(* IEC 61131-3 sources: daoli-st-library/DL_Device (part 13) *)

(* ---- FB_DL_AxisEncBatteryWatch.st ---- *)
(*
    FB_DL_AxisEncBatteryWatch —— 绝对值编码器备用电池欠压监视与预警
    ------------------------------------------------------------------
    组件名称  : FB_DL_AxisEncBatteryWatch
    分类      : DL_Device / AxisHealth
    前缀      : FB_DL_
    版本      : 1.0.0
    溯源      : 借鉴点 —— 设备级粗粒度监视（AOI 粒度族）的「双阈值分型 +
                确认延时 + 锁存预警」组织方式，以及 NE107 健康分级公开条款
                （fault → eMaintenanceReq，warn → eOutOfSpec）。
                本件只借鉴**组织方式与分级语义**，判据 / 阈值 / 码位 100% 自有。
                clean-room 声明 —— 零代码行复制（来源闭源，按最严口径零接触）；
                定时与沿检测仅用 IEC 61131-3 标准库 TON / R_TRIG。
                许可证 —— 本件 MIT；来源标签 t2-6-rockwell-aoi（次源
                t2-8-ne107）仅作语义参考，不包含其任何受版权保护的实现。
    平台      : 纯 IEC 61131-3，CODESYS 3.5 / TwinCAT 3 / InoProShop / Machine Expert 通用
    作者      : 道莅代码库 · PLC编程专家（R71 构建轮 · 批 1 · 序号 3）
    ------------------------------------------------------------------
    功能说明  : 监视绝对值编码器备用电池电压 fBattV，双阈值迟滞判定：
                故障线 fFaultV（低于即电池将尽，断电将丢参考点）与预警线
                fWarnV（低于即建议更换），两线各带独立回差 fHystV 防临界抖振；
                越线须持续 tConfirm 才确认，确认后：
                预警线 → bWarn（实时位）+ bReplaceSoon（**锁存**建议更换位，
                电压回升不清除，必须 bReset 上升沿才解除 —— 电池已劣化属
                事实性结论，瞬时恢复不改判）；
                故障线 → bFault（锁存）+ 故障码。
                非有限电压（断线 / ADC 故障）→ **直接置 bFault 并锁存**
                （电池状态不明比欠压更危险，安全侧收紧，不等确认延时）。
                依赖声明：TYPE E_DL_Ne107Status（属主 I_DL_DeviceHealth.st，
                只引用不重声明，枚举全库唯一定义）；仅 Standard.library
                （TON / R_TRIG / ABS），零厂商方言。
                确认定时器 _tonWarn / _tonFault 每周期无条件调用（规则 ⑦），
                IN 为显式条件（含已确认自保持与回差释放线）。
    错误码    : 16#0002_3770 组态非法（阈值倒置 fWarnV <= fFaultV / 回差为负 /
                            回差吞没线间距 / 阈值非有限 / 幅值超域），锁存 —— 故障级
                16#0002_3771 电池电压非有限（断线 / ADC 故障），直接锁存 —— 故障级
                16#0002_3772 电池欠压越过故障线并经确认（断电将丢参考点），锁存
                            —— 故障级
                16#0002_3773 电池欠压越过预警线并经确认（建议更换）—— 信息级，
                            不置 bError（R45：预警不算故障）
                16#0002_3774 电压越出典型域 [0, 5] V（编码器电池典型域），趋势
                            参考 —— 信息级，不置 bError；不拦截照判（负电压亦
                            必然低于故障线，判定方向天然安全）
    码位总账  : 16#0002_3770 用 ｜ 16#0002_3771 用 ｜ 16#0002_3772 用 ｜
                16#0002_3773 用 ｜ 16#0002_3774 用
    状态机    : N/A —— 单相监视，无顺序状态机，无自有 ENUM / CASE 可写；
                两路确认计时由 TON 实例自持，属定时器状态而非顺序状态；
                健康出口复用既有枚举 E_DL_Ne107Status（只引用）
    边界与披露: 一 组态判据逐项点名（R272）：fWarnV / fFaultV / fHystV 全部
                   纳入非有限闸；阈值倒置（fWarnV <= fFaultV）拦截；
                   fHystV < 0 拦截；fHystV >= (fWarnV - fFaultV) 拦截（回差
                   吞没线间距时两线无迟滞带，判据恒真）；
                二 输入非有限 → 直接故障锁存（不走过闸判定集合，安全侧赋值
                   不引用本闸判定内的量，防自证循环）；
                三 失能（bEn = FALSE）语义写死（R303）：bWarn / bReplaceSoon /
                   bFault 输出全清零、bError 清零、码清零，但 _bFault /
                   _bWarnLatch 锁存位**不被失能清除**（失能是操作态，不是
                   复位），必须 bReset 上升沿才解除 —— 两者语义分离；
                四 定时器 _tonWarn / _tonFault 无论失能 / 故障 / 正常均在段 8
                   无条件调用，IN 为段 7 计算出的显式条件；
                五 阈值默认域标注：编码器备用电池典型域 0~5 V，fWarnV 默认
                   3.0 V / fFaultV 默认 2.7 V 仅为锂-二氧化锰扣式电池组的
                   常见参考值，**不构成工程承诺**，实际阈值以编码器手册为准；
                六 电压越域（0~5 V 外）只报信息级不拦截：判定方向与电压
                   单调性一致（越低越险），越域照判不产生危险侧偏差；
                七 锁存解除路径唯一：bReset 上升沿（R188，可到达、引脚可满足）；
                八 零全局变量、零 VAR_EXTERNAL、零物理地址、零数组下标、无除法。
    分工声明  : FB_DL_BrakeWearAccum（磨损累计）、FB_DL_SpindleWarmupSeq（热机
                顺控）等运动健康件互不相干；本件只做编码器备用电池电压域，
                不消费轴状态、不下发轴指令（R31 运动家族高危区纪律）。
    修订记录  : 2026-11-22 v1.0.0 首次入库（R71 构建轮 · 批 1 · 序号 3）
*)
FUNCTION_BLOCK FB_DL_AxisEncBatteryWatch
VAR_INPUT
    fBattV    : LREAL;                     (* 编码器备用电池电压，[V]，典型域 0..5 / the encoder backup battery voltage *)
    fWarnV    : LREAL := 3.0;              (* 预警阈值，[V]，须 > fFaultV（默认值为参考非承诺）/ the warn threshold, must exceed fFaultV *)
    fFaultV   : LREAL := 2.7;              (* 故障阈值，[V]，须 < fWarnV（默认值为参考非承诺）/ the fault threshold, must be under fWarnV *)
    fHystV    : LREAL := 0.1;              (* 迟滞回差带宽（两线共用独立回差量），[V]，域 [0, fWarnV - fFaultV) / the hysteresis band *)
    tConfirm  : TIME := T#2S;              (* 欠压确认延时，[ms]，须 >= T#0S / the undervoltage confirmation delay *)
    bEn       : BOOL := TRUE;              (* 使能，[标志]，FALSE 时出口清零（R303）/ the enable, FALSE clears the outlets *)
    bReset    : BOOL := FALSE;             (* 故障 / 预警复位，[标志]，上升沿唯一解除 / the reset, its rising edge is the only release *)
END_VAR
VAR_OUTPUT
    bWarn        : BOOL;                   (* 预警实时位（确认成立且未破回差线），[标志] / the live warn flag, confirmed and not released *)
    bFault       : BOOL;                   (* 故障锁存位（故障线确认或电压非有限），[标志] / the latched fault flag *)
    bReplaceSoon : BOOL;                   (* 建议更换锁存位（预警确认后保持至复位），[标志] / the latched replace-soon flag, held until reset *)
    eHealth      : E_DL_Ne107Status;       (* NE107 健康出口（fault → eMaintenanceReq，warn → eOutOfSpec）/ the NE 107 health outlet *)
    bValid       : BOOL;                   (* 出口可用，失能或锁存故障为 FALSE / the outlets usable *)
    bError       : BOOL;                   (* 故障标志，存在锁存故障时为 TRUE / the fault flag, raised while latched *)
    nErrCode     : UDINT;                  (* 错误码，0 = 正常，锁存回放 / the error id, 0 = ok, replayed from the latch *)
END_VAR
VAR
    _rtReset    : R_TRIG;                  (* 复位上升沿检测实例（无条件调用）/ the reset rising edge instance *)
    _tonWarn    : TON;                     (* 预警线确认延时实例（无条件调用）/ the warn line confirmation timer *)
    _tonFault   : TON;                     (* 故障线确认延时实例（无条件调用）/ the fault line confirmation timer *)
    _bFault     : BOOL;                    (* 故障锁存位，仅 bReset 上升沿解除 / the internal latched fault bit *)
    _bWarnLatch : BOOL;                    (* 建议更换锁存位，仅 bReset 上升沿解除 / the internal latched warn bit *)
    _nCodeLatch : UDINT;                   (* 锁存成因码，故障期回放 / the latched cause code, replayed while faulted *)
    _bCfgBad    : BOOL;                    (* 组态非法标志（逐拍重算，仅用于首次锁存）/ the configuration fault flag *)
    _bInBad     : BOOL;                    (* 电压非有限标志（逐拍重算）/ the input fault flag *)
    _bOutDom    : BOOL;                    (* 电压越典型域标志（逐拍重算，仅报信息级）/ the out-of-typical-domain flag *)
    _bRun       : BOOL;                    (* 运行许可 = 使能 且 无锁存故障 / the run permit *)
    _bWarnCond  : BOOL;                    (* 预警确认条件（含自保持与回差，送 TON）/ the warn confirmation condition *)
    _bFaultCond : BOOL;                    (* 故障确认条件（含自保持与回差，送 TON）/ the fault confirmation condition *)
END_VAR

// 段 1｜出口预置（统一出口预置，R256）/ segment 1, preset every outlet
bWarn        := FALSE;                     // 预警实时位预清零 / preset the live warn flag false
bFault       := FALSE;                     // 故障出口预清零 / preset the fault outlet false
bReplaceSoon := FALSE;                     // 建议更换出口预清零 / preset the replace-soon outlet false
eHealth      := E_DL_Ne107Status.eUnknown; // 健康出口预置未知（首拍语义）/ preset the health outlet to unknown
bValid       := FALSE;                     // 可用标志预清零 / preset the valid flag false
bError       := FALSE;                     // 故障标志预清零 / preset the error flag false
nErrCode     := 0;                         // 错误码预置无错 / preset the code to zero
_bWarnCond   := FALSE;                     // 预警条件预清零 / preset the warn condition false
_bFaultCond  := FALSE;                     // 故障条件预清零 / preset the fault condition false

// 段 2｜复位沿检测（无条件调用，规则 ⑦）/ segment 2, the reset edge instance, called unconditionally
_rtReset(CLK := bReset);                   // 每周期无条件刷新 / refreshed every scan without exception

// 段 3｜锁存解除：仅 bReset 上升沿，锁存码同步清零（唯一解除边，R188）/ segment 3, the only latch release edge
IF _rtReset.Q THEN                         // 复位上升沿 / the reset rising edge
    _bFault     := FALSE;                  // 解除故障锁存 / release the fault latch
    _bWarnLatch := FALSE;                  // 解除建议更换锁存 / release the replace-soon latch
    _nCodeLatch := 0;                      // 清锁存码（可到达的清除边）/ clear the latched code, a reachable clearing edge
END_IF

// 段 4｜组态守卫（边界一逐项点名，R272）/ segment 4, the configuration guard
_bCfgBad := (fWarnV <= fFaultV)                                          // 阈值倒置或重合（预警线必须高于故障线）/ the thresholds reversed or coincident
         OR (fHystV < 0.0)                                               // 回差为负 / a negative hysteresis
         OR (fHystV >= (fWarnV - fFaultV))                               // 回差吞没线间距 / the hysteresis swallows the line gap
         OR (fWarnV <> fWarnV) OR ((fWarnV - fWarnV) <> 0.0)             // 预警阈值非有限 / the warn threshold non finite
         OR (fFaultV <> fFaultV) OR ((fFaultV - fFaultV) <> 0.0)         // 故障阈值非有限 / the fault threshold non finite
         OR (fHystV <> fHystV) OR ((fHystV - fHystV) <> 0.0);            // 回差非有限 / the hysteresis non finite

// 段 5｜输入守卫：电压非有限即危险（状态不明 > 欠压，安全侧收紧）/ segment 5, the input guard
_bInBad := (fBattV <> fBattV) OR ((fBattV - fBattV) <> 0.0); // 电压非有限（NaN 自反判 + Inf 差值自反判，R79）/ the voltage non finite
_bOutDom := (fBattV < 0.0) OR (fBattV > 5.0);               // 电压越典型域 [0,5] V（信息级，不拦截照判）/ the voltage out of the typical domain

// 段 6｜首次成因锁存（故障期内不重推断，回放锁存码，R189）/ segment 6, the first-cause latch
IF NOT _bFault THEN                        // 未锁存时才有资格登记成因 / a cause is registered only while not latched
    IF _bCfgBad THEN                       // 组态非法（优先归因，组态是根因）/ an illegal configuration, the root cause first
        _bFault     := TRUE;               // 置故障锁存 / latch the fault
        _nCodeLatch := 16#0002_3770;       // 故障级：组态非法 / fault level: an illegal configuration
    ELSIF _bInBad THEN                     // 电压非有限（状态不明，直接锁存不等延时）/ the voltage non finite, latch at once
        _bFault     := TRUE;               // 置故障锁存 / latch the fault
        _nCodeLatch := 16#0002_3771;       // 故障级：电压非有限 / fault level: a non finite voltage
    END_IF
END_IF

// 段 7｜运行许可与确认条件计算（分支内不调用任何定时器）/ segment 7, the run permit and the conditions
_bRun := bEn AND NOT _bFault;              // 使能且无锁存故障 / enabled and not latched
IF _bRun THEN                              // 运行许可成立 / the run permit holds
    _bWarnCond  := (fBattV < fWarnV) OR (_tonWarn.Q AND NOT (fBattV > (fWarnV + fHystV)));  // 预警条件：破预警线，或已确认且未回升破回差线
    _bFaultCond := (fBattV < fFaultV) OR (_tonFault.Q AND NOT (fBattV > (fFaultV + fHystV))); // 故障条件：破故障线，或已确认且未回升破回差线
    IF _bFaultCond THEN                    // 故障线条件成立（过确认延时后锁存）/ the fault line condition holds
        IF NOT _bFault THEN                // 未锁存才登记 / register only while not latched
            IF _tonFault.Q THEN            // 故障线经确认延时 / the fault line confirmed
                _bFault     := TRUE;       // 置故障锁存 / latch the fault
                _nCodeLatch := 16#0002_3772; // 故障级：欠压越故障线 / fault level: under the fault line
            END_IF
        END_IF
    END_IF
    IF _bWarnCond AND _tonWarn.Q THEN      // 预警线经确认延时 / the warn line confirmed
        _bWarnLatch := TRUE;               // 建议更换锁存（复位才解除，边界三）/ latch the replace-soon flag
    END_IF
ELSE                                       // 失能或锁存故障 / disabled or latched
    _bWarnCond  := FALSE;                  // 条件清零，计时器随之复位 / clear the condition, the timer resets
    _bFaultCond := FALSE;                  // 条件清零 / clear the condition
END_IF

// 段 8｜定时器无条件周期调用（规则 ⑦，IN 为显式条件）/ segment 8, unconditional timer calls
_tonWarn(IN := _bWarnCond, PT := tConfirm);    // 预警确认计时，每周期无条件刷新 / the warn confirmation timer
_tonFault(IN := _bFaultCond, PT := tConfirm);  // 故障确认计时，每周期无条件刷新 / the fault confirmation timer

// 段 9｜出口映射（名实双出口同源，R191）/ segment 9, the outlet mapping
IF _bRun THEN                              // 运行许可成立（无锁存故障）/ the run permit holds, not latched
    bWarn  := _bWarnCond AND _tonWarn.Q;   // 预警实时位：运行中且确认完成 / the live warn flag, confirmed while running
    bFault := FALSE;                       // 无锁存故障，故障出口为假 / no latched fault, the outlet false
    bReplaceSoon := _bWarnLatch;           // 建议更换出口与锁存同源 / the replace-soon outlet shares its latch
    bValid := TRUE;                        // 出口可用 / the outlets usable
    IF bWarn THEN                          // 预警确认成立 / the warn confirmed
        nErrCode := 16#0002_3773;          // 信息级：建议更换（不置 bError，R45）/ info level: replace soon
        eHealth  := E_DL_Ne107Status.eOutOfSpec;   // 预警 → 超出规格 / warn, out of specification
    ELSE                                   // 无预警 / no warn
        eHealth := E_DL_Ne107Status.eOk;   // 正常 / ok
    END_IF
ELSE                                       // 失能或锁存故障（出口清零相）/ disabled or latched, the clearing phase
    IF NOT bEn THEN                        // 失能优先于故障归因（操作态，边界三）/ a disable takes precedence, an operator state
        bWarn   := FALSE;                  // 失能相出口清零（R303）/ zero the outlets while disabled
        bFault  := FALSE;                  // 出口清零（锁存保留）/ the outlet cleared, the latch kept
        bReplaceSoon := FALSE;             // 出口清零（锁存保留）/ the outlet cleared, the latch kept
        bError  := FALSE;                  // 失能不是故障 / a disabled block is not a fault
        nErrCode := 0;                     // 失能不发码 / no code while disabled
        eHealth := E_DL_Ne107Status.eCheckFunction; // 失能 → 功能检查（信号暂无效）/ disabled, function check
    ELSE                                   // 锁存故障相（失能优先级之上）/ the latched fault phase
        bFault  := TRUE;                   // 故障出口与锁存同源 / the fault outlet shares the latch
        bReplaceSoon := _bWarnLatch;       // 建议更换出口与锁存同源 / the replace-soon outlet shares its latch
        bWarn   := FALSE;                  // 故障相预警实时位清零（归并到故障出口）/ the live warn cleared in the fault phase
        bError  := TRUE;                   // 故障标志置位 / raise the fault flag
        nErrCode := _nCodeLatch;           // 回放锁存码 / replay the latched code
        eHealth := E_DL_Ne107Status.eMaintenanceReq; // 故障 → 需要维护 / maintenance required
    END_IF
END_IF
IF _bRun AND (NOT _bFault) AND _bOutDom THEN // 运行中且无锁存故障且越典型域 / running, not latched, out of domain
    IF nErrCode = 0 THEN                   // 不覆盖更高优先级码（信息级让位）/ never overrides a higher priority code
        nErrCode := 16#0002_3774;          // 信息级：电压越典型域 / info level: out of the typical domain
    END_IF
END_IF
END_FUNCTION_BLOCK

(* ---- FB_DL_BcdFieldPanelIO.st ---- *)
(*
  FB_DL_BcdFieldPanelIO  —  面板 BCD 拨码阵列采集/输出 / BCD thumbwheel field panel IO assembly
  分类 Category : DL_Device
  码位 Code     : 16#03_2_17
  段位说明      : 03_2 段低半字节 00~0F 已满（05 为历史空穴留存），R38 已进位 12/13 段，
                  本轮续用 1x 段，本件启用 17 格（R192）
  版本 Version  : 1.0.0
  来源 Source   : t2-1-lgf-converter — BCD 转换族的设备级阵列组装待挖项
  溯源 Origin   : clean-room 实现，未复制任何源码行
                  （与 FC_DL_BcdToWord / FC_DL_WordToBcd 分工：那两件是单路原子，本件是设备级阵列 IO 组装）
  功能 Function : 1) 4 位十进制拨码（16 位输入阵列）逐位消抖（FB_DL_SignalDebounce ×16）；
                  2) 消抖后按 4 bit/位组装 BCD 字 → FC_DL_BcdToWord 逐位解码 → 设定值 uSetValue；
                  3) 位码非法（半字节 > 9）持续 tInvalidTo → 故障级锁存（接线/拨码故障），bReset 解除；
                  4) 稳定值变化沿 bNewValue 单拍脉冲（内部锁存 + 单拍收口，禁同拍抹除）；
                  5) 输出路径：uDisplayVal 经 FC_DL_WordToBcd 回 BCD 字供面板灯显。
  边界 Boundary : ① 16 只消抖实例在主体首部 FOR 循环内无条件刷新（每拍必调，等效无条件域）；
                  ② 位序约定：abDigBits 下标 0 = 个位 BCD bit0，下标 4k..4k+3 = 第 k 位十进制位；
                  ③ tDebounce = T#0S 时消抖直通（消抖件原生语义，透传不钳制）；
                  ④ 组态域闸：tInvalidTo 非正按 1s 兜底（防非法组态令故障永不锁存）；
                  ⑤ 无状态机 CASE 主相（采集型 FB）：故障经锁存位承载，无跨相 TON 复用问题。
  依赖 Depends  : FB_DL_SignalDebounce（实例化 ×16）/ FC_DL_BcdToWord / FC_DL_WordToBcd（函数调用）
  码表 Error codes（本件格 03_2_17，子码步进 +0x100）:
    16#0003_0117 信息级：稳定设定值变化沿已捕获（bNewValue 拍）
    16#0003_0217 故障级：位码非法持续超 tInvalidTo（半字节 > 9，接线/拨码故障），锁存至复位
    16#0003_0317 信息级：回显 BCD 编码饱和（uDisplayVal > 9999，WordToBcd 溢出口径透传）

  修订历史 Revision :
    2026-11-19  v1.0.0  R39 首版（批次 2 · 序号 9）
*)

FUNCTION_BLOCK FB_DL_BcdFieldPanelIO
VAR_INPUT
    abDigBits  : ARRAY[0..15] OF BOOL;    // 拨码原始位输入阵列，下标 0 = 个位 bit0 / Raw digit bit inputs, index 0 = units bit0
    tDebounce  : TIME := T#20MS;          // 逐位消抖延时 [ms]，T#0S = 直通 / Per-bit debounce delay
    tInvalidTo : TIME := T#1S;            // 位码非法持续判据 [ms]，域 > 0（非法组态按 1s 兜底）/ Invalid-code persistence time
    uDisplayVal: UINT := 0;               // 面板回显十进制值 [0..9999]，越限走饱和路径 / Display value for the panel echo
    bReset     : BOOL := FALSE;           // 故障复位，上升沿生效 / Fault reset, rising edge
END_VAR
VAR_OUTPUT
    uSetValue  : UINT;                    // 稳定设定值 [0..9999]（逐位解码合成）/ Stable setpoint value
    bSetValid  : BOOL;                    // 设定值有效（无非法半字节）/ Setpoint validity flag
    anDigVal   : ARRAY[0..3] OF UINT;     // 逐位十进制值 [0..9]（故障位为垃圾值，以 bSetValid 为准）/ Per-digit decimal values
    uBcdEcho   : WORD;                    // 回显 BCD 码字（每半字节一位十进制）/ Echo BCD word for panel lamps
    bNewValue  : BOOL;                    // 稳定设定值变化沿，单拍脉冲 [-] / Stable value change edge, single-cycle pulse
    bError     : BOOL;                    // 故障锁存，仅故障级码置位，bReset 清除 [-] / Fault latch, cleared by reset
    uErrorId   : UDINT;                   // 事件码，0 = 无事件（故障级锁存回放）/ Event code, fault codes latched
END_VAR
VAR
    afbDeb     : ARRAY[0..15] OF FB_DL_SignalDebounce;  // 逐位消抖实例阵列，主体首部无条件刷新 / Per-bit debounce instances
    tonInvalid : TON;                     // 位码非法持续计时（单用途，无跨相复用）/ Invalid-code persistence timer
    rtReset    : R_TRIG;                  // 复位上升沿 / Reset rising edge
    i0         : INT;                     // 位遍历索引 [0..15]，移位量同域严格非负 / Bit loop index, also the shift amount
    _uStable   : WORD;                    // 消抖后稳定 BCD 字 / Debounced stable BCD word
    _uStablePrv: WORD;                    // 上拍稳定 BCD 字（变化沿基准）/ Previous stable BCD word, edge basis
    _bNibBad   : BOOL;                    // 本拍存在非法半字节 / Invalid nibble present this cycle
    _bInit     : BOOL := FALSE;           // 首扫标志，初值 FALSE，判据 NOT bInit（R19 范式）/ First-scan flag
    _bNewLatch : BOOL;                    // 变化沿内部锁存（单拍收口源）/ Change-edge internal latch
    _uEchoErr  : UDINT;                   // WordToBcd 回显错误码透传 / WordToBcd echo error passthrough
    _uDigErr0  : UDINT;                   // 个位 BcdToWord 错误码透传 / Units-digit decode error passthrough
    _uDigErr1  : UDINT;                   // 十位 BcdToWord 错误码透传 / Tens-digit decode error passthrough
    _uDigErr2  : UDINT;                   // 百位 BcdToWord 错误码透传 / Hundreds-digit decode error passthrough
    _uDigErr3  : UDINT;                   // 千位 BcdToWord 错误码透传 / Thousands-digit decode error passthrough
    _uInfo     : UDINT;                   // 本拍信息码，每拍重算 / Transient info code this cycle
    _uFault    : UDINT;                   // 故障码锁存寄存 / Latched fault code register
    _bFault    : BOOL;                    // 故障锁存位 / Latched fault bit
END_VAR
VAR CONSTANT
    DL_BFP_DIG_MASK : WORD := 16#000F;    // 半字节提取掩码（低 4 位）/ Nibble extraction mask
    DL_BFP_INVALID_TO_FBK : TIME := T#1S; // 非法持续判据兜底值 [ms] / Persistence-time fallback value
END_VAR

(* —— 段 0：定时器与边沿实例无条件周期刷新（R7 红线；消抖阵列在 FOR 内每拍全量刷新） —— *)
rtReset(CLK := bReset);                                         // 复位沿刷新，每拍必调
FOR i0 := 0 TO 15 DO                                            // 消抖阵列每拍全量刷新（等效无条件域）
    afbDeb[i0](bRawInput := abDigBits[i0],                      // 原始位输入
               tRiseDelay := tDebounce,                         // 上升确认延时（组态透传）
               tFallDelay := tDebounce,                         // 下降确认延时（组态透传）
               bEnable := TRUE);                                // 消抖恒使能
END_FOR
tonInvalid(IN := _bNibBad, PT := MAX(tInvalidTo, DL_BFP_INVALID_TO_FBK));   // 非法持续计时（单用途，组态兜底）

(* —— 段 1：单拍量预清零（锁存量 _uFault/_bFault/_bNewLatch/_uStablePrv 不入清单，R187①） —— *)
_uInfo := 16#0000_0000;             // 信息码每拍重算
_bNibBad := FALSE;                  // 非法半字节标志预清零
_bNewLatch := FALSE;                // 变化沿锁存预清零（组装段单点置位）
bNewValue := FALSE;                 // 变化沿出口单拍（统一出口映射）
uErrorId := 16#0000_0000;           // 事件码缺省无事件

(* —— 段 2：稳定 BCD 字组装（消抖后位 → 半字节拼接；移位量 = 下标，0..15 严格域内） —— *)
FOR i0 := 0 TO 15 DO
    IF afbDeb[i0].bStable THEN
        _uStable := _uStable OR SHL(WORD#1, i0);    // 置位（移位量归一：下标即移位量，非负）
    ELSE
        _uStable := _uStable AND NOT SHL(WORD#1, i0);   // 清位（移位量同域）
    END_IF
END_FOR

(* —— 段 3：首扫初始化（R19 唯一合法范式） —— *)
IF NOT _bInit THEN
    _uStablePrv := _uStable;        // 首扫：变化沿基准同步为当前稳定字
    _bInit := TRUE;
END_IF

(* —— 段 4：逐位 BCD 解码（FC_DL_BcdToWord 原子 ×4；非法半字节聚合） —— *)
FC_DL_BcdToWord(uBcd := _uStable AND 16#000F, uErrorId => _uDigErr0);   // 个位解码
FC_DL_BcdToWord(uBcd := SHR(_uStable, 4) AND 16#000F, uErrorId => _uDigErr1);   // 十位解码（SHR 正向移位，量归一）
FC_DL_BcdToWord(uBcd := SHR(_uStable, 8) AND 16#000F, uErrorId => _uDigErr2);   // 百位解码
FC_DL_BcdToWord(uBcd := SHR(_uStable, 12) AND 16#000F, uErrorId => _uDigErr3);  // 千位解码
IF (_uDigErr0 <> 0) OR (_uDigErr1 <> 0) OR (_uDigErr2 <> 0) OR (_uDigErr3 <> 0) THEN
    _bNibBad := TRUE;               // 本拍存在非法半字节（任一位 > 9）
END_IF
anDigVal[0] := FC_DL_BcdToWord(uBcd := _uStable AND 16#000F);           // 个位值（错误路径返回 0，安全侧）
anDigVal[1] := FC_DL_BcdToWord(uBcd := SHR(_uStable, 4) AND 16#000F);   // 十位值
anDigVal[2] := FC_DL_BcdToWord(uBcd := SHR(_uStable, 8) AND 16#000F);   // 百位值
anDigVal[3] := FC_DL_BcdToWord(uBcd := SHR(_uStable, 12) AND 16#000F);  // 千位值
uSetValue := anDigVal[0] + anDigVal[1] * 10 + anDigVal[2] * 100 + anDigVal[3] * 1000;   // 十进制合成

(* —— 段 5：故障锁存（非法持续到点才锁存，瞬时切换不误报） —— *)
IF tonInvalid.Q THEN
    _uFault := 16#0003_0217;        // 故障级：位码非法持续超限
    _bFault := TRUE;
END_IF
IF rtReset.Q THEN
    _bFault := FALSE;               // 清故障锁存位（唯一解除路径：bReset 上升沿）
    _uFault := 16#0000_0000;
END_IF

(* —— 段 6：有效性出口与变化沿（内部锁存 → 统一出口单拍，两段式收口） —— *)
bSetValid := NOT _bNibBad;          // 有效性 = 本拍无非法半字节（瞬时口径）
IF (NOT _bNibBad) AND (_uStable <> _uStablePrv) THEN
    _bNewLatch := TRUE;             // 稳定字变化：内部锁存置位（段 1 已预清零，同拍不抹）
    _uInfo := 16#0003_0117;         // 信息级：变化沿已捕获
END_IF
_uStablePrv := _uStable;            // 变化沿基准更新（段尾单点）
bNewValue := _bNewLatch;            // 出口 = 内部锁存（置位同拍不被抹）

(* —— 段 7：回显 BCD 编码（FC_DL_WordToBcd 原子，越限饱和码透传） —— *)
uBcdEcho := FC_DL_WordToBcd(uVal := uDisplayVal, uErrorId => _uEchoErr);
IF _uEchoErr <> 0 THEN
    _uInfo := 16#0003_0317;         // 信息级：回显饱和（覆盖变化沿码，回显状态优先）
END_IF

(* —— 段 8：事件码单点回放（故障锁存优先） —— *)
IF _bFault THEN
    uErrorId := _uFault;            // 故障锁存码回放
    bError := TRUE;
ELSE
    uErrorId := _uInfo;             // 信息码
    bError := FALSE;
END_IF

END_FUNCTION_BLOCK

(* ---- FB_DL_BilletShearGaugeSeq.st ---- *)
(*
  Component : FB_DL_BilletShearGaugeSeq
  Category  : DL_Device
  Type      : FB
  Complexity: C2
  VERSION   : v1.0.0
  功能      : 铸锭定尺剪切时序控制：ENUM 八态（Idle/Feed/Measure/Clamp/Shear/Trim/Release/Fault），按定尺长度送进、夹紧确认后剪切，首件去头尾。
  开源溯源  : 道莅原创 clean-room 自研（无外部代码引用）｜License: MIT
  边界条件  : ① 定尺长度须 > 1e-9、各段时长为 0 判组态非法，拒绝启动并锁存故障；
              ② 首件定尺 = 定尺长度 + 去头尾长度，去头尾仅首件执行一次；
              ③ 夹紧超时 / 松开超时均判故障，故障锁存唯一解除路径 = bReset 上升沿。
*)

TYPE E_DL_ShearPhase :
(
    eIdle    := 0,    (* 空闲：等启动沿 / Idle waiting start edge *)
    eFeed    := 10,   (* 送进：至定尺到位 / Feeding to gauge length *)
    eMeasure := 20,   (* 测长：稳定驻留 / Measuring dwell *)
    eClamp   := 30,   (* 夹紧：至夹紧反馈 / Clamping to feedback *)
    eShear   := 40,   (* 剪切：剪切保持 / Shearing hold *)
    eTrim    := 50,   (* 去头尾：首件端部切除 / Head-trim cut on first piece *)
    eRelease := 60,   (* 松开：至松开确认 / Releasing to confirmation *)
    eFault   := 90    (* 故障：锁存待复位 / Fault latched *)
);
END_TYPE

FUNCTION_BLOCK FB_DL_BilletShearGaugeSeq
VAR_INPUT
    bEnable     : BOOL;   (* 使能电平 [-] Enable level *)
    bReset      : BOOL;   (* 复位上升沿，清故障锁存 [-] Reset edge *)
    bStart      : BOOL;   (* 启动上升沿 [-] Start edge *)
    fLengthMm   : REAL;   (* 送进实测长度 [mm] Measured feed length *)
    fGaugeLenMm : REAL;   (* 定尺长度 [mm] Gauge length setpoint *)
    fTrimLenMm  : REAL;   (* 去头尾长度 [mm] Head trim length *)
    bClampFb    : BOOL;   (* 夹紧到位反馈 [-] Clamp feedback *)
    bShearFb    : BOOL;   (* 剪切到位反馈 [-] Shear feedback *)
    tMeasure    : TIME;   (* 测长驻留 [ms] Measuring dwell *)
    tShear      : TIME;   (* 剪切保持 [ms] Shear hold *)
    tTrim       : TIME;   (* 去头尾保持 [ms] Trim hold *)
    tClampTo    : TIME;   (* 夹紧超时 [ms] Clamp timeout *)
    tReleaseTo  : TIME;   (* 松开超时 [ms] Release timeout *)
END_VAR
VAR_OUTPUT
    bFeedRun    : BOOL;              (* 送进运行输出 [-] Feed run output *)
    bClampCmd   : BOOL;              (* 夹紧指令输出 [-] Clamp command *)
    bShearCmd   : BOOL;              (* 剪切指令输出 [-] Shear command *)
    bTrimCmd    : BOOL;              (* 去头尾刀指令输出 [-] Trim cut command *)
    bReleaseCmd : BOOL;              (* 松开指令输出 [-] Release command *)
    nPieceCnt   : INT;               (* 完成件数 [-] Finished piece counter *)
    ePhase      : E_DL_ShearPhase;   (* 相位出口，段尾单点映射 [-] Phase outlet *)
    bError      : BOOL;              (* 故障锁存标志 [-] Fault latch flag *)
    uErrId      : UDINT;             (* 事件码，0 = 无事件 [-] Event code *)
END_VAR
VAR
    rtReset   : R_TRIG;   (* 复位沿实例，每拍无条件刷新 / Reset edge *)
    rtStart   : R_TRIG;   (* 启动沿实例，每拍无条件刷新 / Start edge *)
    tonMeasure: TON;      (* 测长驻留计时（独立实例） / Measuring timer *)
    tonShear  : TON;      (* 剪切保持计时（独立实例） / Shear timer *)
    tonTrim   : TON;      (* 去头尾保持计时（独立实例） / Trim timer *)
    tonClampTo: TON;      (* 夹紧超时（专用超时件） / Clamp timeout *)
    tonRelTo  : TON;      (* 松开超时（专用超时件） / Release timeout *)
    _ePhase   : E_DL_ShearPhase := E_DL_ShearPhase.eIdle;  (* 内部相位 / Internal phase *)
    _bFault   : BOOL;     (* 故障锁存位（锁存量） / Latched fault bit *)
    _uFault   : UDINT;    (* 故障码锁存（锁存量） / Latched fault code *)
    _bFirst   : BOOL;     (* 首件标志（锁存量） / First piece flag *)
    _bCfgBad  : BOOL;     (* 组态非法当拍量 [-] Config illegal flag *)
    _bNonFin  : BOOL;     (* 输入非有限当拍量 [-] Non-finite input flag *)
    fTargetMm : REAL;     (* 本件定尺目标 [mm] Target length of this piece *)
END_VAR
VAR CONSTANT
    DL_EPS : REAL := 1.0E-9;   (* 浮点比较容差 [无量纲] Float compare tolerance *)
    DL_ZERO: REAL := 0.0;      (* 零常量 [-] Zero constant *)
END_VAR

(* —— 段 0｜沿与定时器每拍无条件刷新（禁置于 IF/CASE 内，使能挂 IN 引脚） —— *)
rtReset(CLK := bReset);
rtStart(CLK := bStart);
tonMeasure(IN := (_ePhase = E_DL_ShearPhase.eMeasure) AND (NOT _bFault), PT := tMeasure);
tonShear  (IN := (_ePhase = E_DL_ShearPhase.eShear)   AND (NOT _bFault), PT := tShear);
tonTrim   (IN := (_ePhase = E_DL_ShearPhase.eTrim)    AND (NOT _bFault), PT := tTrim);
tonClampTo(IN := (_ePhase = E_DL_ShearPhase.eClamp)   AND (NOT _bFault), PT := tClampTo);
tonRelTo  (IN := (_ePhase = E_DL_ShearPhase.eRelease) AND (NOT _bFault), PT := tReleaseTo);

(* —— 段 1｜每拍量预清零（锁存量 _bFault/_uFault/_bFirst/nPieceCnt 不入清单） —— *)
uErrId := 16#0000_0000;
_bCfgBad := FALSE;
_bNonFin := FALSE;

(* —— 段 2｜复位沿：故障一次性清干净，相位回空闲，首件标志复原 —— *)
IF rtReset.Q THEN
    _bFault := FALSE;
    _uFault := 16#0000_0000;
    _bFirst := TRUE;
    _ePhase := E_DL_ShearPhase.eIdle;
END_IF

(* —— 段 3｜组态闸与非有限判据（覆盖定尺长度与各段时长） —— *)
IF (fGaugeLenMm <= DL_EPS) OR (fTrimLenMm < DL_ZERO) OR (tMeasure = T#0S)
   OR (tShear = T#0S) OR (tTrim = T#0S) OR (tClampTo = T#0S) OR (tReleaseTo = T#0S) THEN
    _bCfgBad := TRUE;
END_IF
IF (fLengthMm <> fLengthMm) OR ((fLengthMm - fLengthMm) <> 0.0)
   OR (fGaugeLenMm <> fGaugeLenMm) OR ((fGaugeLenMm - fGaugeLenMm) <> 0.0)
   OR (fTrimLenMm <> fTrimLenMm) OR ((fTrimLenMm - fTrimLenMm) <> 0.0) THEN
    _bNonFin := TRUE;
END_IF

(* —— 段 4｜本件定尺目标：首件叠加去头尾长度 —— *)
IF _bFirst THEN
    fTargetMm := fGaugeLenMm + fTrimLenMm;
ELSE
    fTargetMm := fGaugeLenMm;
END_IF

(* —— 段 5｜主状态机：八态全覆盖 + ELSE 兜底 —— *)
CASE _ePhase OF
E_DL_ShearPhase.eIdle:
    bFeedRun := FALSE; bClampCmd := FALSE; bShearCmd := FALSE;
    bTrimCmd := FALSE; bReleaseCmd := FALSE;
    IF rtStart.Q AND bEnable AND (NOT _bFault) AND (NOT _bCfgBad) AND (NOT _bNonFin) THEN
        nPieceCnt := 0;
        _bFirst := TRUE;
        _ePhase := E_DL_ShearPhase.eFeed;
    ELSIF rtStart.Q AND (_bFault OR _bCfgBad OR _bNonFin) THEN
        _bFault := TRUE;                  (* 带病启动拒绝 / Reject start with bad config *)
        _uFault := 16#0024_0001;
        _ePhase := E_DL_ShearPhase.eFault;
    END_IF

E_DL_ShearPhase.eFeed:
    bFeedRun := TRUE; bClampCmd := FALSE; bShearCmd := FALSE;
    bTrimCmd := FALSE; bReleaseCmd := FALSE;
    IF _bNonFin THEN
        _bFault := TRUE; _uFault := 16#0024_0002;   (* 故障级：长度反馈非有限 *)
        _ePhase := E_DL_ShearPhase.eFault;
    ELSIF fLengthMm >= fTargetMm THEN
        _ePhase := E_DL_ShearPhase.eMeasure;        (* 迁出条件 1：定尺到位 *)
    ELSIF NOT bEnable THEN
        _ePhase := E_DL_ShearPhase.eIdle;           (* 迁出条件 2：使能撤销回安全态 *)
    END_IF

E_DL_ShearPhase.eMeasure:
    bFeedRun := FALSE; bClampCmd := FALSE; bShearCmd := FALSE;
    bTrimCmd := FALSE; bReleaseCmd := FALSE;
    IF tonMeasure.Q THEN
        _ePhase := E_DL_ShearPhase.eClamp;          (* 迁出条件 1：测长驻留完成 *)
    ELSIF NOT bEnable THEN
        _ePhase := E_DL_ShearPhase.eIdle;           (* 迁出条件 2：使能撤销 *)
    END_IF

E_DL_ShearPhase.eClamp:
    bFeedRun := FALSE; bClampCmd := TRUE; bShearCmd := FALSE;
    bTrimCmd := FALSE; bReleaseCmd := FALSE;
    IF bClampFb THEN
        _ePhase := E_DL_ShearPhase.eShear;          (* 迁出条件 1：夹紧反馈到位 *)
    ELSIF tonClampTo.Q THEN
        _bFault := TRUE; _uFault := 16#0024_0003;   (* 故障级：夹紧超时 *)
        _ePhase := E_DL_ShearPhase.eFault;
    END_IF

E_DL_ShearPhase.eShear:
    bFeedRun := FALSE; bClampCmd := TRUE; bShearCmd := TRUE;
    bTrimCmd := FALSE; bReleaseCmd := FALSE;
    IF bShearFb OR tonShear.Q THEN
        IF _bFirst THEN
            _ePhase := E_DL_ShearPhase.eTrim;       (* 首件：追加去头尾刀 *)
        ELSE
            _ePhase := E_DL_ShearPhase.eRelease;    (* 迁出条件 1：剪切到位或保持到时 *)
        END_IF
    ELSIF NOT bEnable THEN
        _ePhase := E_DL_ShearPhase.eIdle;           (* 迁出条件 2：使能撤销 *)
    END_IF

E_DL_ShearPhase.eTrim:
    bFeedRun := FALSE; bClampCmd := TRUE; bShearCmd := FALSE;
    bTrimCmd := TRUE; bReleaseCmd := FALSE;
    IF tonTrim.Q THEN
        _ePhase := E_DL_ShearPhase.eRelease;        (* 迁出条件 1：去头尾保持完成 *)
    ELSIF NOT bEnable THEN
        _ePhase := E_DL_ShearPhase.eIdle;           (* 迁出条件 2：使能撤销 *)
    END_IF

E_DL_ShearPhase.eRelease:
    bFeedRun := FALSE; bClampCmd := FALSE; bShearCmd := FALSE;
    bTrimCmd := FALSE; bReleaseCmd := TRUE;
    IF NOT bClampFb THEN
        nPieceCnt := nPieceCnt + 1;                 (* 完成件数累加：仅在迁出拍执行一次 *)
        _bFirst := FALSE;                           (* 首件完成，后续按纯定尺 *)
        _ePhase := E_DL_ShearPhase.eFeed;           (* 迁出条件 1：松开确认到位 *)
    ELSIF tonRelTo.Q THEN
        _bFault := TRUE; _uFault := 16#0024_0004;   (* 故障级：松开超时 *)
        _ePhase := E_DL_ShearPhase.eFault;
    END_IF

E_DL_ShearPhase.eFault:
    bFeedRun := FALSE; bClampCmd := FALSE; bShearCmd := FALSE;
    bTrimCmd := FALSE; bReleaseCmd := FALSE;        (* 故障相：全部输出走安全侧 *)

ELSE
    _bFault := TRUE;                                (* 兜底：非法相位锁存 *)
    _uFault := 16#0024_0009;
    _ePhase := E_DL_ShearPhase.eFault;
END_CASE

(* —— 段 6｜相位与故障码出口单点映射 —— *)
ePhase := _ePhase;
bError := _bFault;
IF _bFault AND (_uFault <> 16#0000_0000) THEN
    uErrId := _uFault;                              (* 故障码锁存回放 / Latched fault replay *)
END_IF
END_FUNCTION_BLOCK

(* ---- FB_DL_BmsPdiGateway.st ---- *)
(*
  FB_DL_BmsPdiGateway  —  楼宇侧 PDI 对象网关轮询（调度 + 异常上报） / Building-side PDI object gateway polling: scheduling plus exception report
  分类 Category : DL_Device
  版本 Version  : 1.0.0
  来源 Source   : t1-4-codesys-forge — 网关轮询族零检索深化（与 PdiReadScheduler 调度底座分工：那件为底层调度，本件为楼宇网关应用件）
  溯源 Origin   : clean-room 实现，未复制任何源码行
  功能 Function : 1) 轮询调度：bPollTick 调用方节拍沿驱动，对象索引 0..uObjCnt-1
                  轮转（uObjCnt 域闸 1..8），每拍采信当前对象 bPollOk / fObjVal
                  契约快照，逐对象连续失败计数 auFailCnt；
                  2) 异常上报：连续失败达 uFailTo → 0528 首出对象锁存
                  （nFirstFailObj 记首出号，R190 归因唯一）；对象值非有限
                  → 0529 防御锁存（NaN 自反判）；
                  3) 成功承载：失败计数清零 + 值快照写入 afObjVal + 信息级
                  042E；首出锁存拍发 042F；
                  4) 故障级：0528 对象连续失败超阈 / 0529 对象值非有限 /
                  052A 组态非法（对象数越域）+ ELSE 兜底归并；
                  5) 信息级三码：轮询成功 / 超时上报 / 网关复位（单拍沿）；
                  6) 解除式全当拍量（R240 落地），逐 BOOL 标注见段 4。
  边界 Boundary : ① 分段理由（R192）：段 0003 故障带 03A0~03FF 于 R42 用尽，
                  启用 05xx 副带续编，避开 0590~0599 判错位段；
                  ② 组态闸：uObjCnt = 0 或 > 8 或 uFailTo = 0 → 052A 锁存，
                  轮询停发；对象索引域 0..7 由 uObjCnt 域闸与常量 8 结构性限定；
                  ③ 失败计数 USINT 饱和前置判（防回绕）；
                  ④ 无 GVL 依赖：纯引脚输入输出，无外部变量引用，无物理 IO 地址。
  依赖 Depends  : Standard.library（R_TRIG）
  码表 Error codes（Device 段 0003，窗口 0528~052A / 042E~0430）:
    16#0003_0528 故障级：对象连续失败超阈锁存（首出对象号入 nFirstFailObj），锁存至 bReset
    16#0003_0529 故障级：对象值非有限锁存（防御兜底），锁存至 bReset
    16#0003_052A 故障级：组态非法（对象数/失败阈域非法）或相位落 ELSE 兜底（归并声明），锁存至 bReset
    16#0003_042E 信息级：轮询成功沿（对象值快照写入拍）
    16#0003_042F 信息级：超时上报沿（首出锁存拍）
    16#0003_0430 信息级：网关复位沿（台账清零拍）
  修订历史 Revision :
    2026-11-19  v1.0.0  R42 首版（批次 4 · 序号 5）
*)

TYPE E_DL_BpgState :
(
    eIdle  := 0,     // 未使能：不轮询 / Idle, not polling
    ePoll  := 10,    // 轮询中：逐对象承载 / Poll, per-object engaged
    eFault := 90     // 故障：首出或非有限锁定 / Fault, latched
);
END_TYPE

FUNCTION_BLOCK FB_DL_BmsPdiGateway
VAR_INPUT
    bPollTick    : BOOL := FALSE;     // 轮询节拍沿（调用方驱动）[-] / Poll tick edge from caller
    bPollOk      : BOOL := FALSE;     // 当前对象轮询成功（当拍量契约）[-] / Current-object poll success
    fObjVal      : REAL := 0.0;       // 当前对象值 [工程单位]，bPollOk 当拍采信 / Current-object value
    uObjCnt      : USINT := 8;        // 对象总数 [1..8]，域闸 / Object count
    uFailTo      : USINT := 3;        // 连续失败阈 [次]，域 > 0 / Consecutive-fail threshold
    bGwEn        : BOOL := FALSE;     // 网关使能（电平）[-] / Gateway enable, level
    bReset       : BOOL := FALSE;     // 复位，上升沿清故障锁存与台账 / Reset edge
END_VAR
VAR_OUTPUT
    eState       : E_DL_BpgState;     // 状态出口，段尾单点映射 / State outlet
    nObjIdx      : DINT;              // 当前轮询对象号 [0..7]，-1 = 未轮询 / Current polling object index
    afObjVal     : ARRAY[0..7] OF REAL;   // 逐对象值快照 [工程单位] / Per-object value snapshots
    auFailCnt    : ARRAY[0..7] OF USINT;  // 逐对象连续失败计数 [次] / Per-object fail counts
    nFirstFailObj: DINT;              // 首出失败对象号 [0..7]，-1 = 无首出 / First failed object index
    bError       : BOOL;              // 故障锁存标志 / Fault latch flag
    nErrId       : UDINT;             // 事件码，0 = 无事件 / Event code
END_VAR
VAR
    rtPollTick   : R_TRIG;            // 轮询节拍沿实例，无条件刷新 / Poll tick edge instance
    rtReset      : R_TRIG;            // 复位沿实例，无条件刷新 / Reset edge instance
    _eState      : E_DL_BpgState := E_DL_BpgState.eIdle;  // 内部相位（CASE 唯一写入目标）/ Internal phase
    _nObjCursor  : UDINT := 0;        // 轮转游标 [0..uObjCnt-1] / Round-robin cursor
    _nIdx        : DINT;              // 阵列循环索引 [-] / Array loop index
    _bValNonFin  : BOOL;              // 对象值非有限当拍量 [-] / Object-value non-finite flag
    _bFault      : BOOL;              // 故障锁存位（锁存量）/ Latched fault bit
    _uFault      : UDINT;             // 故障码锁存（锁存量）/ Latched fault code
    _uInfo       : UDINT;             // 信息码，每拍重算 / Transient info code
END_VAR

(* —— 段 0：沿实例无条件周期刷新（禁置于 IF/CASE 内） —— *)
_bValNonFin := (fObjVal <> fObjVal)
            OR ((fObjVal - fObjVal) <> (fObjVal - fObjVal));    // 值非有限防御（NaN 自反 + 差值自减）
rtPollTick(CLK := bPollTick);       // 轮询节拍沿（每拍必调）
rtReset(CLK := bReset);             // 复位沿（每拍必调）

(* —— 段 1：单拍量预清零（锁存量 _bFault/_uFault 与计数阵列不入清单，禁同拍抹除） —— *)
_uInfo := 16#0000_0000;             // 信息码每拍重算
nObjIdx := -1;                      // 对象号缺省 -1
nErrId := 16#0000_0000;             // 事件码缺省无事件

(* —— 段 2：复位沿 + 组态域闸（判据当拍量） —— *)
IF rtReset.Q THEN                   // rtReset.Q = 当拍量
    _bFault := FALSE;               // 清故障锁存位
    _uFault := 16#0000_0000;        // 清故障锁存码
    nFirstFailObj := -1;            // 首出对象号恢复哨兵
    FOR _nIdx := 0 TO 7 DO          // 台账逐对象清零
        auFailCnt[_nIdx] := 0;      // 失败计数清零
        afObjVal[_nIdx] := 0.0;     // 值快照清零
    END_FOR
    _uInfo := 16#0003_0430;         // 信息级：网关复位沿
END_IF
IF (uObjCnt < 1) OR (uObjCnt > 8) OR (uFailTo = 0) THEN      // 域闸（1..8 与失败阈）
    _uFault := 16#0003_052A;        // 故障级：组态非法
    _bFault := TRUE;                // 故障标志与码位配对（R45）
END_IF

(* —— 段 3：轮询沿承载（判据当拍量；对象索引由域闸 1..8 结构性限域） —— *)
IF rtPollTick.Q AND (_eState = E_DL_BpgState.ePoll) AND (NOT _bFault) THEN
    _nObjCursor := (_nObjCursor + 1) MOD UDINT(uObjCnt);    // 轮转游标（模基数域闸 > 0，无除零）
    nObjIdx := UDINT_TO_DINT(_nObjCursor);          // 当前对象号（域 0..uObjCnt-1 ⊆ 0..7）
    IF bPollOk THEN                 // 成功承载（当拍量契约）
        auFailCnt[nObjIdx] := 0;    // 失败计数清零
        IF NOT _bValNonFin THEN     // 值快照仅非有限闸通过后写入（FB32-7 保持槽闸）
            afObjVal[nObjIdx] := fObjVal;       // 值快照写入
        END_IF
        _uInfo := 16#0003_042E;     // 信息级：轮询成功沿
    ELSE                            // 失败承载
        IF auFailCnt[nObjIdx] < 255 THEN
            auFailCnt[nObjIdx] := auFailCnt[nObjIdx] + 1;   // 计数递增（饱和前置判防回绕）
        END_IF
        IF (auFailCnt[nObjIdx] >= uFailTo) AND (nFirstFailObj = -1) THEN
            nFirstFailObj := nObjIdx;   // 首出对象号锁定（仅首个写入）
            _uFault := 16#0003_0528;    // 故障级：连续失败超阈
            _bFault := TRUE;
            _uInfo := 16#0003_042F;     // 信息级：超时上报沿
        END_IF
    END_IF
    IF _bValNonFin AND bPollOk THEN // 成功契约但值非有限：防御锁存（0529 独立归因）
        _uFault := 16#0003_0529;    // 故障级：对象值非有限
        _bFault := TRUE;
    END_IF
END_IF

(* —— 段 4：故障解除式（R240 落地，逐 BOOL 标注）：
     rtReset.Q = 当拍量；bPollOk = 当拍量；NOT bGwEn = 当拍量。
     均不含锁存量（_bFault/_uFault），解除边真实可达（轮询恢复 + 撤使能 + 复位沿）。 —— *)
IF rtReset.Q AND bPollOk AND (NOT bGwEn) THEN
    _bFault := FALSE;               // 清故障锁存位（锁存量，仅此当拍量解除沿可清）
    _uFault := 16#0000_0000;        // 清故障锁存码（锁存量，仅本当拍量解除沿可清）
    IF _eState = E_DL_BpgState.eFault THEN
        _eState := E_DL_BpgState.eIdle;     // 故障相迁出：回未使能
    END_IF
END_IF

(* —— 段 5：相位机（CASE 全覆盖 + ELSE 兜底） —— *)
CASE _eState OF

E_DL_BpgState.eIdle:
    IF bGwEn AND (NOT _bFault) THEN
        _eState := E_DL_BpgState.ePoll;     // 使能：进轮询相
    END_IF

E_DL_BpgState.ePoll:
    IF (NOT _bFault) AND (NOT bGwEn) THEN
        _eState := E_DL_BpgState.eIdle;     // 撤使能：回未使能相
    END_IF
    (* 首出/非有限迁出在段 3 承载（置 _bFault 后次拍迁故障相） *)

E_DL_BpgState.eFault:
    ;                               // 故障相：轮询冻结，等解除沿（段 4 承载迁出）

ELSE
    _uFault := 16#0003_052A;        // 故障级：非法相位兜底（归并组态码，码表声明）
    _bFault := TRUE;
    _eState := E_DL_BpgState.eFault;    // 强制回故障相

END_CASE

(* —— 段 6：出口单点映射（名实同源；锁存码回放，禁同拍抹除） —— *)
IF _bFault THEN
    nErrId := _uFault;              // 故障锁存码回放
    nObjIdx := -1;                  // 故障相对象号恢复未轮询哨兵
ELSE
    nErrId := _uInfo;               // 信息码
END_IF
bError := _bFault;                  // 故障标志与锁存位同源
eState := _eState;                  // 状态出口单点映射

END_FUNCTION_BLOCK

(* ---- FB_DL_BoilerFlueCondenseGuard.st ---- *)
(*
  FB_DL_BoilerFlueCondenseGuard  —  锅炉烟气冷凝防护（排烟温度低限联锁 + 回水温度钳制） / Boiler flue-gas condensation guard with low flue-temperature interlock and return-water clamping
  分类 Category : DL_Device
  版本 Version  : 1.0.0
  来源 Source   : t1-2-oscat-building — 楼宇锅炉防冷凝保护族深化
  溯源 Origin   : 道莅 clean-room 实现；排烟温度低限联锁 + 回水温度低限钳制为公开锅炉防低温腐蚀保护逻辑，未复制任何源码行
  功能 Function : 1) 三级判据：排烟温度 fFlueTempC 低于报警限 fFlueLoC → 冷凝风险信息位；
                  低于联锁限 fFlueLoLoC 且持续 tConfirm → 联锁撤销燃烧器许可；
                  2) 回水温度钳制：fReturnTempC 低于 fReturnMinC 时输出 bReturnClamp 请求（提高回水），
                  仅在燃烧器许可有效时给出；
                  3) 故障级单码 052C / 信息级 0432 = 冷凝风险进入沿（由无风险转风险单拍）。
  接口 Interface: 输入排烟温度/两级限值/回水温度/回水下限/确认延时；输出许可与风险位
  边界 Boundary : ① 组态闸：fFlueLoLoC >= fFlueLoC（联锁限须低于报警限）、fFlueLoC <= 0.0、
                  fReturnMinC < 0.0、tConfirm <= T#0S → 052C 锁存；
                  ② 温度非有限（NaN 自反 + Inf 差值自减）→ 052C 锁存，燃烧器许可撤销（安全侧）；
                  ③ 低限判据为「<=」单侧直比（限值语义明确，无容差歧义），回水钳制同为单侧直比；
                  ④ 一个 TON + 两个 R_TRIG 段 0 无条件调用；⑤ 故障相迁出唯一路径 = bReset 上升沿；
                  ⑥ 零全局耦合：无 GVL / VAR_EXTERNAL / %I %Q %M 直接地址。
  依赖 Depends  : Standard.library（TON / R_TRIG）
  码表 Error codes（Device 分段见下，故障窗口 052C / 信息窗口 0432）:
    16#0003_052C 故障级：烟气冷凝防护故障总码（组态非法 / 温度非有限），锁存至 bReset 上升沿；
                 归因见 eCause，不新增码位（派单硬约束单码）
    16#0003_0432 信息级：冷凝风险进入沿（无风险 → 风险，单拍）
    分段理由：段 0003 故障带 03A0~03FF 于 R42 用尽，启用 05xx 副带续编，避开 0590~0599 判错位段。
  修订历史 Revision :
    2026-11-19  v1.0.0  R43 首版（批次 4 · 序号 16）
*)

TYPE E_DL_BfgState :
(
    eIdle     := 0,   // 未使能：许可撤销 / Idle, permit withdrawn
    eGuard    := 10,  // 防护监视中（许可有效） / Guarding with permit valid
    eLockout  := 20,  // 联锁动作（许可撤销） / Interlocked, permit withdrawn
    eFault    := 90   // 故障锁存相 / Fault latched phase
);
END_TYPE

TYPE E_DL_BfgCause :
(
    eNone       := 0, // 无故障成因 / No cause
    eCfgIllegal := 1, // 组态非法 / Illegal configuration
    eNonFinite  := 2  // 温度非有限 / Non-finite temperature
);
END_TYPE

FUNCTION_BLOCK FB_DL_BoilerFlueCondenseGuard
VAR_INPUT
    fFlueTempC   : REAL := 0.0;        // 排烟温度 [°C] / Flue gas temperature
    fFlueLoC     : REAL := 90.0;       // 冷凝风险报警限 [°C]，域 > 0 / Condensation alarm limit
    fFlueLoLoC   : REAL := 70.0;       // 联锁限 [°C]，须低于报警限 / Interlock limit
    fReturnTempC : REAL := 0.0;        // 回水温度 [°C] / Return water temperature
    fReturnMinC  : REAL := 55.0;       // 回水温度下限 [°C]，域 >= 0 / Return water minimum
    tConfirm     : TIME := T#30S;      // 联锁确认延时 [ms]，域 > 0 / Interlock confirmation delay
    bEnable      : BOOL := FALSE;      // 防护使能（电平）[-] / Guard enable
    bReset       : BOOL := FALSE;      // 复位命令，上升沿清故障 [-] / Reset edge
END_VAR
VAR_OUTPUT
    eState       : E_DL_BfgState;      // 状态出口，段 6 单点映射 / State outlet
    eCause       : E_DL_BfgCause;      // 故障成因出口（R190） / Fault cause outlet
    bBurnerPermit: BOOL;               // 燃烧器许可 [-] / Burner permit
    bCondenseRisk: BOOL;               // 冷凝风险位 [-] / Condensation risk flag
    bReturnClamp : BOOL;               // 回水温度钳制请求 [-] / Return-water clamping request
    bError       : BOOL;               // 故障锁存标志 [-] / Fault latch flag
    nErrId       : UDINT;              // 事件码，0 = 无事件 / Event code
END_VAR
VAR
    _eState      : E_DL_BfgState := E_DL_BfgState.eIdle;   // 内部相位（CASE 唯一写入目标） / Internal phase
    _eCause      : E_DL_BfgCause := E_DL_BfgCause.eNone;   // 故障成因锁存（锁存量） / Latched cause
    tonConfirm   : TON;                // 联锁确认计时，每周期无条件调用 / Confirmation timer
    rtReset      : R_TRIG;             // 复位沿实例，每周期无条件调用 / Reset edge
    rtRisk       : R_TRIG;             // 风险沿实例，每周期无条件调用 / Risk edge
    _bRisk       : BOOL;               // 冷凝风险当拍量 [-] / Risk verdict
    _bLoLo       : BOOL;               // 低于联锁限当拍量 [-] / Below interlock limit
    _bRetLow     : BOOL;               // 回水低于下限当拍量 [-] / Return water below minimum
    _bNonFin     : BOOL;               // 温度非有限当拍量 [-] / Non-finite temperature
    _bCfgBad     : BOOL;               // 组态非法当拍量 [-] / Config illegal
    _bFault      : BOOL;               // 故障锁存位（锁存量） / Latched fault bit
    _uFault      : UDINT;              // 故障码锁存（锁存量） / Latched fault code
    _uInfo       : UDINT;              // 信息码，每拍重算 / Transient info code
END_VAR

(* —— 段 0：沿实例与定时器无条件周期刷新 + 当拍量判据 —— *)
_bRisk := fFlueTempC <= fFlueLoC;                                            // 冷凝风险（单侧直比） / Risk verdict
_bLoLo := fFlueTempC <= fFlueLoLoC;                                          // 低于联锁限 / Below interlock
_bRetLow := fReturnTempC < fReturnMinC;                                      // 回水低于下限 / Return below minimum
_bNonFin := (fFlueTempC <> fFlueTempC) OR (fReturnTempC <> fReturnTempC)
         OR ((fFlueTempC - fFlueTempC) <> (fFlueTempC - fFlueTempC))
         OR ((fReturnTempC - fReturnTempC) <> (fReturnTempC - fReturnTempC));  // NaN 自反 + Inf 差值自减 / NaN and Inf
_bCfgBad := (fFlueLoLoC >= fFlueLoC) OR (fFlueLoC <= 0.0) OR (fReturnMinC < 0.0)
            OR (tConfirm <= T#0S);                                           // 组态非法当拍量 / Config illegal
rtReset(CLK := bReset);                                                      // 复位沿，每拍必调 / Reset edge
rtRisk(CLK := _bRisk AND (NOT _bFault));                                     // 风险沿（故障相屏蔽） / Risk edge
tonConfirm(IN := (_eState = E_DL_BfgState.eGuard) AND _bLoLo, PT := tConfirm);   // 联锁确认计时 / Interlock timer

(* —— 段 1：单拍量预清零（锁存量不入清单） —— *)
_uInfo := 16#0000_0000;            // 信息码每拍重算 / Info recomputed
bBurnerPermit := FALSE;            // 许可缺省撤销（安全侧缺省） / Permit default withdrawn
bCondenseRisk := FALSE;            // 风险位缺省 FALSE / Risk default
bReturnClamp := FALSE;             // 钳制请求缺省 FALSE / Clamp default
nErrId := 16#0000_0000;            // 事件码缺省无事件 / Event code default

(* —— 段 2：复位沿 + 组态域闸 —— *)
IF rtReset.Q THEN                              // rtReset.Q = 当拍量 / current scan
    _bFault := FALSE;                          // 清故障锁存位（锁存量） / Clear fault latch
    _uFault := 16#0000_0000;                   // 清故障锁存码（锁存量） / Clear fault code
    _eCause := E_DL_BfgCause.eNone;            // 清成因（锁存量） / Clear cause
    IF _eState = E_DL_BfgState.eFault THEN
        _eState := E_DL_BfgState.eIdle;        // 故障相迁出：回未使能 / Fault exit to idle
    END_IF
    IF _eState = E_DL_BfgState.eLockout THEN
        _eState := E_DL_BfgState.eGuard;       // 联锁相复位迁出：回防护（恢复许可） / Lockout exit to guard
    END_IF
END_IF
IF _bCfgBad THEN                               // 组态域闸 / Config gate
    _uFault := 16#0003_052C;                   // 故障级：防护故障总码（05xx 副带） / Device fault code
    _eCause := E_DL_BfgCause.eCfgIllegal;      // 归因：组态非法 / Cause: illegal config
    _bFault := TRUE;                           // 标志与码位配对（R45） / Flag paired with code
END_IF
IF (NOT _bFault) AND _bNonFin THEN             // 非有限锁存 / Non-finite latch
    _uFault := 16#0003_052C;
    _eCause := E_DL_BfgCause.eNonFinite;       // 归因：非有限 / Cause: non-finite
    _bFault := TRUE;
END_IF

(* —— 段 3：联锁确认（低于联锁限持续 tConfirm 即进联锁相） —— *)
IF (NOT _bFault) AND (_eState = E_DL_BfgState.eGuard) AND tonConfirm.Q THEN
    _eState := E_DL_BfgState.eLockout;         // 进联锁相（许可撤销） / Enter lockout
END_IF

(* —— 段 4：故障解除式（R240；全当拍量）：rtReset.Q / NOT _bCfgBad / NOT _bNonFin —— *)
IF rtReset.Q AND (NOT _bCfgBad) AND (NOT _bNonFin) THEN
    _bFault := FALSE;                          // 清故障锁存位（锁存量） / Clear fault latch
    _uFault := 16#0000_0000;                   // 清故障锁存码（锁存量） / Clear fault code
    _eCause := E_DL_BfgCause.eNone;            // 清成因（锁存量） / Clear cause
END_IF

(* —— 段 4A：故障锁存相位迁移闸 —— *)
IF _bFault AND (_eState <> E_DL_BfgState.eFault) THEN
    _eState := E_DL_BfgState.eFault;           // 锁存即入故障相 / Latch enters fault phase
END_IF

(* —— 段 5：相位机（CASE 全覆盖 + ELSE 兜底） —— *)
CASE _eState OF

E_DL_BfgState.eIdle:
    IF bEnable AND (NOT _bFault) THEN          // 使能条件 / Enable gate
        _eState := E_DL_BfgState.eGuard;       // 进防护相 / Enter guard
    END_IF

E_DL_BfgState.eGuard:
    bBurnerPermit := NOT _bLoLo;               // 许可：未低于联锁限即允许 / Permit unless below interlock
    bCondenseRisk := _bRisk;                   // 风险位（相内按当拍量给出） / Risk flag
    bReturnClamp := _bRetLow AND bBurnerPermit; // 回水钳制请求（许可有效时） / Return clamp request
    IF rtRisk.Q THEN                           // 风险进入沿 / Risk entrance edge
        _uInfo := 16#0003_0432;                // 信息级：冷凝风险进入沿 / Info: risk entrance
    END_IF
    IF NOT bEnable THEN                        // 撤使能：许可撤销，回未使能 / Disable withdraws permit
        _eState := E_DL_BfgState.eIdle;
    ELSIF NOT _bRisk THEN                      // 风险消失：保持防护相（不迁移） / Risk cleared, stay
        ;
    END_IF

E_DL_BfgState.eLockout:
    bBurnerPermit := FALSE;                    // 联锁相：许可强制撤销 / Permit forced withdrawn
    bCondenseRisk := TRUE;                     // 联锁相风险位恒真 / Risk latched high
    IF NOT _bLoLo THEN                         // 排烟温度回到联锁限之上（事件） / Flue temperature recovered
        _eState := E_DL_BfgState.eGuard;       // 恢复防护相 / Back to guard
    ELSIF NOT bEnable THEN                     // 撤使能：回未使能 / Disable returns idle
        _eState := E_DL_BfgState.eIdle;
    END_IF

E_DL_BfgState.eFault:
    ;                                          // 故障相：许可撤销，仅段 4 复位沿可迁出 / Permit withdrawn, reset only

ELSE
    _uFault := 16#0003_052C;                   // 故障级：非法相位兜底（归并总码） / Illegal phase fallback
    _eCause := E_DL_BfgCause.eCfgIllegal;      // 归因：相位非法归并组态 / Cause: phase illegal
    _bFault := TRUE;
    _eState := E_DL_BfgState.eFault;           // 强制回故障相 / Force fault phase

END_CASE

(* —— 段 6：出口单点映射（名实同源；故障相许可强制撤销） —— *)
IF _bFault THEN
    bBurnerPermit := FALSE;                    // 故障相许可强制撤销（安全侧） / Permit forced withdrawn
    bReturnClamp := FALSE;                     // 故障相钳制请求强制 FALSE / Clamp forced false
    nErrId := _uFault;                         // 故障锁存码回放 / Replay latched code
ELSE
    nErrId := _uInfo;                          // 信息码 / Transient info
END_IF
bError := _bFault;                             // 故障标志同源 / Flag from latch
eState := _eState;                             // 状态出口 / State outlet
eCause := _eCause;                             // 成因出口 / Cause outlet

END_FUNCTION_BLOCK

(* ---- FB_DL_BoothExhaustDamperSeq.st ---- *)
(*
  Name: FB_DL_BoothExhaustDamperSeq
  Category: DL_Device
  Version: 1.0.0
  Round: R89 / 2026-11-25
  开源溯源：clean-room 自研（族 涂装喷涂线，ST 开源生态实测 0 命中，无外部代码引入）
  功能：喷房排风风门开度顺序：起机预吹→生产→清洗大风量→停机，斜坡按周期步进，含卡涩监视。
  边界条件：① 四浮点入参全部过非有限闸；配置越域进冻结分支：输出保持末值 + xValid = FALSE（R191）；
            ② 目标开度按模式赋值：预吹取 min(60 %, 外部设定)、生产取外部设定、清洗取 100 %（大风量）；
            ③ 斜坡步长 = fRampPctPerS × fCycleS，周期非法取 10 ms 缺省；开度钳 0~100 %；
            ④ 卡涩监视：实际开度与斜坡输出偏差 > 10 % 时锁故障（风门卡滞/执行器失气）；
            ⑤ 故障解除唯一路径：故障相内 xStart 释放（R152），清锁存回 eIdle。
  状态机：eIdle / eRamp / eHold / eFault（CASE 含 ELSE 兜底；模式亦用 ENUM + CASE 兜底）。
*)
TYPE E_DL_BedMode :
(
    ePurge   := 0,      (* 预吹模式：低开度预吹 / Purge mode, low opening *)
    eProduce := 1,      (* 生产模式：按外部设定 / Production mode, external setpoint *)
    eClean   := 2       (* 清洗模式：大风量满开 / Cleaning mode, full opening *)
);
END_TYPE
TYPE E_DL_BedsPhase :
(
    eIdle  := 0,        (* 停机相：斜坡回 0 / Stopped, ramping to zero *)
    eRamp  := 10,       (* 斜坡相：向目标开度推进 / Ramping to setpoint *)
    eHold  := 20,       (* 保持相：已在目标开度带内 / Holding at setpoint *)
    eFault := 90        (* 故障相：锁存待释放 / Fault latched, awaiting release *)
);
END_TYPE

FUNCTION_BLOCK FB_DL_BoothExhaustDamperSeq
VAR_INPUT
    xStart : BOOL;              (* 起机命令 [-] Start command *)
    eMode : E_DL_BedMode;       (* 运行模式（0 预吹 / 1 生产 / 2 清洗） [-] Operating mode *)
    fDamperActPct : REAL;       (* 风门实际开度 [%] Damper actual opening [%] *)
    fDamperSpPct : REAL;        (* 生产模式开度设定 [%] Production setpoint opening [%] *)
    fRampPctPerS : REAL;        (* 斜坡速率 [%/s] Ramp rate [%/s] *)
    fCycleS : REAL;             (* 扫描周期 [s] Scan cycle [s] *)
END_VAR
VAR_OUTPUT
    xDamperCmd : BOOL;          (* 风门开命令 [-] Damper open command *)
    fDamperOutPct : REAL;       (* 风门开度输出（斜坡后） [%] Damper opening output [%] *)
    eState : E_DL_BedsPhase;     (* 当前相 [-] Present phase *)
    xValid : BOOL;              (* 配置与链路有效 [-] Configuration and chain valid *)
END_VAR
VAR
    _eState : E_DL_BedsPhase := E_DL_BedsPhase.eIdle;  (* 内部相（CASE 唯一写入目标） [-] Internal phase *)
    _bFaultLatch : BOOL := FALSE;   (* 故障锁存位 [-] Fault latch *)
    _bCfgBad : BOOL := FALSE;       (* 配置非法当拍量 [-] Configuration bad *)
    _bCalcOk : BOOL := FALSE;       (* 本拍计算有效 [-] Calculation valid this scan *)
    _bStuck : BOOL := FALSE;        (* 卡涩判据 [-] Damper stuck *)
    _fOut : REAL := 0.0;            (* 开度斜坡保持量 [%] Opening hold [%] *)
    _fSp : REAL := 0.0;             (* 当拍目标开度 [%] Target opening [%] *)
    _fStep : REAL := 0.0;           (* 单拍斜坡步长 [%] Ramp step [%] *)
    _fCy : REAL := 0.01;            (* 当拍有效周期 [s] Effective cycle [s] *)
END_VAR
VAR CONSTANT
    DL_BDS_EPS : REAL := 1.0E-9;        (* 判据容差 [-] Criterion tolerance *)
    DL_BDS_PURGE : REAL := 60.0;        (* 预吹开度 [%] Purge opening [%] *)
    DL_BDS_CLEAN : REAL := 100.0;       (* 清洗开度 [%] Cleaning opening [%] *)
    DL_BDS_TOL : REAL := 1.0;           (* 到位带半宽 [%] In-position band [%] *)
    DL_BDS_STUCK : REAL := 10.0;        (* 卡涩偏差门限 [%] Stuck deviation threshold [%] *)
    DL_BDS_CYDEF : REAL := 0.01;        (* 缺省扫描周期 [s] Default scan cycle [s] *)
    DL_BDS_PCT_MAX : REAL := 100.0;     (* 开度满量程 [%] Opening full scale [%] *)
END_VAR
(* 非有限闸（NaN 自反 + Inf 差值自减）+ 组态域闸：四浮点入参全枚举（R272） *)
_bCfgBad := (fDamperActPct <> fDamperActPct) OR ((fDamperActPct - fDamperActPct) <> 0.0)
         OR (fDamperSpPct <> fDamperSpPct) OR ((fDamperSpPct - fDamperSpPct) <> 0.0)
         OR (fRampPctPerS <> fRampPctPerS) OR ((fRampPctPerS - fRampPctPerS) <> 0.0)
         OR (fCycleS <> fCycleS) OR ((fCycleS - fCycleS) <> 0.0)
         OR (fDamperActPct < 0.0) OR (fDamperActPct > DL_BDS_PCT_MAX)
         OR (fDamperSpPct < 0.0) OR (fDamperSpPct > DL_BDS_PCT_MAX)
         OR (fRampPctPerS < 1.0) OR (fRampPctPerS > 200.0);
(* 周期派生：非法周期取 10 ms 缺省 *)
IF (fCycleS > 0.0) AND (fCycleS <= 1.0) THEN
    _fCy := fCycleS;
ELSE
    _fCy := DL_BDS_CYDEF;
END_IF
_bCalcOk := xStart AND (NOT _bCfgBad);
(* 目标开度：按模式取值（ENUM + CASE，含 ELSE 兜底） *)
CASE eMode OF
E_DL_BedMode.ePurge:
    IF fDamperSpPct < DL_BDS_PURGE THEN
        _fSp := fDamperSpPct;               (* 预吹取设定与 60 % 的较小者 / Lower of setpoint and 60 % *)
    ELSE
        _fSp := DL_BDS_PURGE;
    END_IF
E_DL_BedMode.eProduce:
    _fSp := fDamperSpPct;                   (* 生产按外部设定 / Production uses setpoint *)
E_DL_BedMode.eClean:
    _fSp := DL_BDS_CLEAN;                   (* 清洗满开 / Cleaning full open *)
ELSE
    _fSp := 0.0;                            (* 非法模式：目标归零 / Illegal mode, zero target *)
END_CASE
(* 停机即目标归零（安全侧） *)
IF NOT _bCalcOk THEN
    _fSp := 0.0;
END_IF
(* 斜坡推进：步长 = 速率 × 周期，方向按目标与当前比较 *)
_fStep := fRampPctPerS * _fCy;
(* 非有限/越界步长闸：NOT(x>=0) 对 NaN 为真，防 NaN 直穿 _fOut 出口 *)
IF NOT ((_fStep >= 0.0) AND (_fStep <= 100.0)) THEN
    _fStep := 0.0;                          (* 步长归零，风门保持原位 / Zero step, hold position *)
END_IF
IF _fOut < (_fSp - DL_BDS_TOL) THEN
    _fOut := _fOut + _fStep;
    IF _fOut > _fSp THEN
        _fOut := _fSp;                      (* 上钳 / Upper clamp *)
    END_IF
ELSIF _fOut > (_fSp + DL_BDS_TOL) THEN
    _fOut := _fOut - _fStep;
    IF _fOut < _fSp THEN
        _fOut := _fSp;                      (* 下钳 / Lower clamp *)
    END_IF
END_IF
(* 卡涩判据：指令与实际偏差超门限（仅在斜坡/保持相监视） *)
_bStuck := ABS(_fOut - fDamperActPct) > DL_BDS_STUCK;
(* 状态机（ENUM + CASE，ELSE 兜底） *)
CASE _eState OF
E_DL_BedsPhase.eIdle:
    IF _bCalcOk THEN
        _eState := E_DL_BedsPhase.eRamp;     (* 起机 → 斜坡 / Start, ramp *)
    END_IF
E_DL_BedsPhase.eRamp:
    IF _bStuck THEN
        _eState := E_DL_BedsPhase.eFault;    (* 卡涩 → 故障 / Stuck, fault *)
    ELSIF ABS(_fOut - _fSp) <= DL_BDS_TOL THEN
        _eState := E_DL_BedsPhase.eHold;     (* 到位 → 保持 / In position, hold *)
    END_IF
E_DL_BedsPhase.eHold:
    IF NOT _bCalcOk THEN
        _eState := E_DL_BedsPhase.eIdle;     (* 停机 → 回斜坡关风门 / Stop, close damper *)
    ELSIF _bStuck THEN
        _eState := E_DL_BedsPhase.eFault;    (* 卡涩 → 故障 / Stuck, fault *)
    ELSIF ABS(_fOut - _fSp) > DL_BDS_TOL THEN
        _eState := E_DL_BedsPhase.eRamp;     (* 目标变化 → 回斜坡 / Target changed, re-ramp *)
    END_IF
E_DL_BedsPhase.eFault:
    _bFaultLatch := TRUE;                   (* 故障相锁存（码由相位表达） / Latch in fault phase *)
    IF NOT xStart THEN
        _bFaultLatch := FALSE;              (* 解除路径：启动释放（R152） / Released by start drop *)
        _eState := E_DL_BedsPhase.eIdle;     (* 回待机 / Back to idle *)
    END_IF
ELSE
    _bFaultLatch := TRUE;                   (* 非法相兜底 / Illegal phase fallback *)
    _eState := E_DL_BedsPhase.eFault;
END_CASE
(* 统一出口（单点赋值）：停机相也照实输出斜坡值，避免风门瞬断 *)
xDamperCmd := (_fOut > 0.5) OR (_eState = E_DL_BedsPhase.eRamp) OR (_eState = E_DL_BedsPhase.eHold);
fDamperOutPct := _fOut;
eState := _eState;
xValid := _bCalcOk;
END_FUNCTION_BLOCK

(* ---- FB_DL_BrakeResistorThermal.st ---- *)
(*
  Name        : FB_DL_BrakeResistorThermal
  Category    : DL_Device
  Version     : 1.0.1
  Purpose     : 变频器制动电阻热累积估算：按 I²·R 瞬时功率逐拍积分成能量，叠加一阶冷却（时间常数 tau）折算温升与能量百分比，给出过载/预警与降额建议；/ Estimate braking-resistor thermal accumulation by integrating I2R power with first-order cooling, yielding temperature rise, energy percentage, overload warnings and a derating hint
  溯源        : 借 t2-6-rockwell-aoi 的分类/参数域组织，clean-room 实现
  Boundary    : ① 组态闸：额定电流/电阻/时间常数/周期/温升额度任一非正 → 锁存故障；
                ② 除零前置：热容/时间常数、能量上限、温升额度的除子均在组态闸保证非按零后使用；
                ③ 非有限电流/温度输入该拍不积分（保留上拍累积值，防污染积分器）；
                ④ 能量百分比饱和 0..100 且过载判据用 >= 阈值直比（阈值来自组态，非浮点等值比较）；
                ⑤ 本件为估算模型，不替代硬件热保护（安全回路须由变频器/热继电器实现）。
  修订记录    : 2026-11-20 v1.0.1：温升改热阻功率比口径（fRiseRated × P/P_rated，R52-09）；组态闸追加能量额度一致性校验（fEnergyMax > I²R·τ 派生上界即故障）并把默认 fEnergyMax 收口为 6000 kJ 派生值；_fPct 饱和处回夹 _fAccJ/_fAccKj 能量上界（R52-10）；eIdle 补 fEnergyPct/fDeratePct 出口镜像并按 dT/dt = -T/tauCool 冷却衰减。
*)
TYPE E_DL_BrtState :
(
    eIdle  := 0,                             (* 未使能 / Disabled *)
    eEst   := 10,                            (* 热累积估算 / Thermal estimation *)
    eFault := 90                             (* 故障锁存相 / Fault latched *)
);
END_TYPE

TYPE E_DL_BrtCause :
(
    eNone       := 0,                        (* 无故障成因 / No cause *)
    eCfgIllegal := 1,                        (* 组态非法：电气参数/时间常数越域 / Illegal config *)
    ePhaseBad   := 2                         (* 非法相位兜底 / Illegal phase fallback *)
);
END_TYPE

FUNCTION_BLOCK FB_DL_BrakeResistorThermal
VAR_INPUT
    fBrakeCurrent : REAL := 0.0;             (* 制动电流实测（RMS），域 >= 0 [A] / Measured braking current RMS *)
    fRatedCurrent : REAL := 20.0;            (* 电阻额定电流，域 > 0 [A] / Rated current, > 0 *)
    fResistance   : REAL := 50.0;            (* 电阻阻值（冷态），域 > 0 [Ohm] / Resistance, > 0 *)
    tCycle        : TIME := T#10MS;          (* 估算周期，域 > T#0S [ms] / Estimation period, > 0 *)
    fTauCool      : REAL := 300.0;           (* 冷却时间常数 tau，域 > 0 [s] / Cooling time constant, > 0 *)
    fEnergyMax    : REAL := 6000.0;          (* 允许累计能量上限（= 可吸收能量，默认为 I²R·τ 派生量 20²·50·300/1000，须 <= 派生上界）[kJ] / Allowed energy budget, <= I2R*tau derived cap *)
    fTempAmb      : REAL := 40.0;            (* 环境温度 [°C] / Ambient temperature *)
    fRiseRated    : REAL := 250.0;           (* 满载（额定）稳态温升，域 > 0 [K] / Steady rise at rated load, > 0 *)
    bEnable       : BOOL := TRUE;            (* 估算使能 [-] / Enable *)
    bReset        : BOOL := FALSE;           (* 复位命令，上升沿清累积能量与故障 [-] / Reset command *)
END_VAR
VAR_OUTPUT
    fEnergyKj    : REAL;                     (* 当前累积能量（净额，含冷却扣除）[kJ] / Accumulated net energy *)
    fEnergyPct   : REAL;                     (* 能量占额度百分比 0..100（饱和）[%] / Energy percentage, saturated *)
    fTempRise    : REAL;                     (* 估算温升（相对环境）[K] / Estimated temperature rise *)
    fTempEst     : REAL;                     (* 估算电阻温度 = 环境 + 温升 [°C] / Estimated resistor temperature *)
    fDeratePct   : REAL;                     (* 降额建议（100 = 不降额，50 = 半载），0..100 [%] / Derating hint, 0..100 *)
    bWarn        : BOOL;                     (* 预警：能量百分比 >= 80% [-] / Warning at 80 percent *)
    bOverload    : BOOL;                     (* 过载：能量百分比 >= 100% [-] / Overload at 100 percent *)
    eState       : E_DL_BrtState;            (* 状态出口 / State outlet *)
    eCause       : E_DL_BrtCause;            (* 故障成因出口（R190 归因唯一） / Fault cause outlet *)
    bError       : BOOL;                     (* 故障锁存标志 [-] / Fault latch flag *)
END_VAR
VAR
    _eState   : E_DL_BrtState := E_DL_BrtState.eIdle;    (* 内部相位（CASE 唯一写入目标） / Internal phase *)
    _eCause   : E_DL_BrtCause := E_DL_BrtCause.eNone;    (* 故障成因锁存量 / Latched cause *)
    rtReset   : R_TRIG;                      (* 复位沿实例，段 0 无条件调用 / Reset edge instance *)
    _bFault   : BOOL;                        (* 故障锁存位 / Latched fault bit *)
    _bCfgBad  : BOOL;                        (* 组态非法当拍量 / Illegal config this scan *)
    _bFinite  : BOOL;                        (* 输入有限性当拍量 / Input finiteness *)
    _fDtSec   : REAL;                        (* 周期折算秒值，域 > eps [s] / Period in seconds *)
    _fPowerW  : REAL;                        (* 本拍制动功率 P = I²·R [W] / Braking power this scan *)
    _fEinJ    : REAL;                        (* 本拍注入能量 [J] / Injected energy this scan *)
    _fEoutJ   : REAL;                        (* 本拍冷却带走能量（一阶）[J] / Energy removed by cooling *)
    _fAccJ    : REAL;                        (* 累积能量内部量（焦耳口径）[J] / Accumulated energy in joules *)
    _fAccKj   : REAL;                        (* 累积能量换算 kJ 中间量 [kJ] / Accumulated energy in kJ *)
    _fPct     : REAL;                        (* 未饱和百分比 [%] / Unclamped percentage *)
    _fRiseEst : REAL;                        (* 温升估算中间量 [K] / Rise estimate intermediate *)
    _fDerate  : REAL;                        (* 降额中间量 [%] / Derate intermediate *)
    _fBudgetKj: REAL;                        (* 能量额度物理上界 I²R·τ 派生量（kJ 口径）[kJ] / Physics energy cap I2R*tau *)
    _fEfullJ  : REAL;                        (* 能量额度满值焦耳换算中间量（回夹用）[J] / Budget in joules for clamping *)
END_VAR
VAR CONSTANT
    DL_BRT_EPS   : REAL := 1.0E-6;           (* 判零容差（REAL 量级）[-] / Epsilon *)
    DL_BRT_J2KJ  : REAL := 1000.0;           (* 焦耳→千焦换算因子（常量除子）[-] / Joules to kJ factor *)
    DL_BRT_PCTMAX: REAL := 100.0;            (* 百分比满量程 [%] / Percentage full scale *)
    DL_BRT_WARN  : REAL := 80.0;             (* 预警门槛 [%] / Warning threshold *)
END_VAR

(* —— 段 0：当拍判据派生 + 实例无条件刷新（R228A） —— *)
_fDtSec := TIME_TO_LREAL(tCycle) / 1000.0;                                     (* 周期秒化（除子常量 1000） / Period to seconds *)
_fBudgetKj := fRatedCurrent * fRatedCurrent * fResistance * fTauCool / DL_BRT_J2KJ;   (* 能量额度物理上界 = I²R·τ（稳态能量平衡，除子为常量）[kJ] / Physics cap I2R*tau *)
_fEfullJ := fEnergyMax * DL_BRT_J2KJ;                                          (* 能量额度满值焦耳换算（回夹上界）[J] / Budget in joules *)
_bCfgBad := NOT (tCycle > T#0S)                                                (* 周期正域闸 / Period gate *)
            OR (fRatedCurrent <= DL_BRT_EPS) OR (fResistance <= DL_BRT_EPS)    (* 电气参数正域闸 / Electrical gates *)
            OR (fTauCool <= DL_BRT_EPS) OR (fEnergyMax <= DL_BRT_EPS)          (* 冷却常数/能量额度正域闸（除零前置） / Cooling and budget gates *)
            OR (fRiseRated <= DL_BRT_EPS)                                      (* 温升额度正域闸 / Rise gate *)
            OR ((fTauCool > DL_BRT_EPS) AND (fEnergyMax > _fBudgetKj));        (* 能量额度一致性校验：应 ≈ I²R·τ 派生量（除子先过正域闸，v1.0.1）/ Budget consistency gate *)
rtReset(CLK := bReset);                                                        (* 复位沿每拍必调 / Reset edge every scan *)
_bFinite := (fBrakeCurrent = fBrakeCurrent) AND (fTempAmb = fTempAmb)          (* NaN 自反闸 / NaN reflex gates *)
            AND ((fBrakeCurrent - fBrakeCurrent) = (fBrakeCurrent - fBrakeCurrent));   (* Inf 差判闸 / Inf gate *)

(* —— 段 1：单拍量预清零（R107） —— *)
bWarn := FALSE;                                                                (* 预警位预清 / Warn preset *)
bOverload := FALSE;                                                            (* 过载位预清 / Overload preset *)

(* —— 段 2：复位沿处理（作用域：清故障 + 清累积能量 + 清出口 + 迁 eIdle，R283 逐项声明） —— *)
IF rtReset.Q THEN
    _bFault := FALSE;                                                          (* 清故障锁存 / Clear fault *)
    _eCause := E_DL_BrtCause.eNone;                                            (* 清成因 / Clear cause *)
    _fAccJ := 0.0;                                                             (* 清累积能量（焦耳） / Clear accumulated joules *)
    fEnergyKj := 0.0;                                                          (* 清能量出口 / Clear energy outlet *)
    fEnergyPct := 0.0;                                                         (* 清百分比出口 / Clear percentage *)
    fTempRise := 0.0;                                                          (* 清温升出口 / Clear rise outlet *)
    fTempEst := fTempAmb;                                                      (* 温度回环境值 / Temperature back to ambient *)
    fDeratePct := DL_BRT_PCTMAX;                                               (* 降额建议回 100%（不降额） / Derate back to 100 *)
    _eState := E_DL_BrtState.eIdle;                                            (* 迁未使能相 / Back to idle *)
END_IF

(* —— 段 3：组态故障锁存（锁存至复位沿，R189） —— *)
IF _bCfgBad AND NOT _bFault THEN
    _bFault := TRUE;                                                           (* 锁存故障位 / Latch fault *)
    _eCause := E_DL_BrtCause.eCfgIllegal;                                      (* 成因：组态非法 / Cause: illegal config *)
    _eState := E_DL_BrtState.eFault;                                           (* 同步迁故障相 / Migrate to fault *)
END_IF

(* —— 段 4：CASE 主状态机（ELSE 兜底迁 eFault，红线 6） —— *)
CASE _eState OF
    E_DL_BrtState.eIdle:                                                       (* 未使能：停机冷却 + 出口镜像 / Disabled: cooling and mirrors *)
        _fAccJ := _fAccJ - (_fAccJ / fTauCool) * _fDtSec;                      (* 停机即按 dT/dt = -T/tauCool 一阶冷却衰减（除子 tau 已过组态闸，v1.0.1） / First-order cooling while idle *)
        IF _fAccJ < 0.0 THEN
            _fAccJ := 0.0;                                                     (* 冷却下限 0：不允许负累积 / Energy floor zero *)
        END_IF
        _fAccKj := _fAccJ / DL_BRT_J2KJ;                                       (* 焦耳→千焦（除子为常量）[kJ] / Joules to kJ *)
        fEnergyKj := _fAccKj;                                                  (* 能量出口镜像 / Energy outlet mirror *)
        _fPct := _fAccKj / fEnergyMax * DL_BRT_PCTMAX;                         (* 占额度百分比：除子额度已过闸 [%] / Percentage of budget *)
        IF _fPct > DL_BRT_PCTMAX THEN
            _fPct := DL_BRT_PCTMAX;                                            (* 上限饱和 100 [%] / Upper saturation *)
        ELSIF _fPct < 0.0 THEN
            _fPct := 0.0;                                                      (* 下限饱和 0 [%] / Lower saturation *)
        END_IF
        fEnergyPct := _fPct;                                                   (* 百分比出口镜像（v1.0.1 补） / Percentage outlet mirror *)
        _fDerate := DL_BRT_PCTMAX - _fPct;                                     (* 降额镜像：能量越满降额越深 [%] / Derate mirror *)
        IF _fDerate < 0.0 THEN
            _fDerate := 0.0;                                                   (* 降额下限 0 / Derate floor *)
        END_IF
        fDeratePct := _fDerate;                                                (* 降额出口镜像（v1.0.1 补） / Derate outlet mirror *)
        fTempRise := 0.0;                                                      (* 无估算语义：温升 0 / No estimation: rise 0 *)
        fTempEst := fTempAmb;                                                  (* 温度 = 环境 / Temperature = ambient *)
        IF bEnable AND NOT _bFault THEN
            _eState := E_DL_BrtState.eEst;                                     (* 使能进入估算 / Enter estimation *)
        END_IF
    E_DL_BrtState.eEst:                                                        (* 估算相：I²R 积分 + 一阶冷却 / Estimation *)
        IF NOT bEnable THEN
            _eState := E_DL_BrtState.eIdle;                                    (* 失能回未使能 / Back to idle *)
        ELSIF _bFinite AND (_fDtSec > DL_BRT_EPS) THEN
            _fPowerW := fBrakeCurrent * fBrakeCurrent * fResistance;            (* 瞬时制动功率 I²·R [W]（乘性，无除零） / Instantaneous I2R power *)
            _fEinJ := _fPowerW * _fDtSec;                                      (* 本拍注入能量 [J] / Injected energy *)
            _fEoutJ := (_fAccJ / fTauCool) * _fDtSec;                          (* 一阶冷却带走能量（除子 tau 已过闸）[J] / First-order cooling *)
            _fAccJ := _fAccJ + _fEinJ - _fEoutJ;                               (* 净额积分（单点写入，无双向双计） / Net integration, single write *)
            IF _fAccJ < 0.0 THEN
                _fAccJ := 0.0;                                                 (* 能量下限 0：不允许负累积 / Energy floor zero *)
            END_IF
            _fAccKj := _fAccJ / DL_BRT_J2KJ;                                   (* 焦耳→千焦 [kJ] / Joules to kJ *)
            fEnergyKj := _fAccKj;                                              (* 能量出口 / Energy outlet *)
            _fPct := _fAccKj / fEnergyMax * DL_BRT_PCTMAX;                     (* 占额度百分比：除子额度已过闸 [%] / Percentage of budget *)
            IF _fPct > DL_BRT_PCTMAX THEN
                _fPct := DL_BRT_PCTMAX;                                        (* 上限饱和 100 [%] / Upper saturation *)
                _fAccJ := _fEfullJ;                                            (* 能量上界回夹 = 额度满值（饱和处同步，v1.0.1，R52-10） / Clamp energy to budget *)
                _fAccKj := fEnergyMax;                                         (* kJ 镜像同步回夹 / Mirror clamp in kJ *)
                fEnergyKj := _fAccKj;                                          (* 能量出口同步回夹 / Energy outlet sync *)
            ELSIF _fPct < 0.0 THEN
                _fPct := 0.0;                                                  (* 下限饱和 0 [%] / Lower saturation *)
            END_IF
            fEnergyPct := _fPct;                                               (* 百分比出口 / Percentage outlet *)
            _fRiseEst := fRiseRated * (_fPowerW / (fRatedCurrent * fRatedCurrent * fResistance));   (* 温升 = 满载稳态温升 × 瞬时功率/额定功率比（热阻口径，除子由组态闸保证 > 0，v1.0.1） / Rise = rated rise times power ratio *)
            IF _fRiseEst < 0.0 THEN
                _fRiseEst := 0.0;                                              (* 温升下限 0 [K] / Rise floor *)
            END_IF
            fTempRise := _fRiseEst;                                            (* 温升出口 [K] / Rise outlet *)
            fTempEst := fTempAmb + _fRiseEst;                                  (* 电阻温度 = 环境 + 温升 [°C] / Estimated temperature *)
            _fDerate := DL_BRT_PCTMAX - _fPct;                                 (* 降额建议：能量越满降额越深 [%] / Derate hint *)
            IF _fDerate < 0.0 THEN
                _fDerate := 0.0;                                               (* 降额下限 0（已过载即全禁） / Derate floor *)
            END_IF
            fDeratePct := _fDerate;                                            (* 降额出口 / Derate outlet *)
            IF _fPct >= DL_BRT_PCTMAX THEN
                bOverload := TRUE;                                             (* 过载：能量额度耗尽 / Overload: budget exhausted *)
            ELSIF _fPct >= DL_BRT_WARN THEN
                bWarn := TRUE;                                                 (* 预警：能量额度达 80% / Warning at 80 percent *)
            END_IF
        END_IF                                                                 (* 非有限输入：不积分，保持上拍累积（边界③） / Non-finite: hold *)
    E_DL_BrtState.eFault:                                                      (* 故障相：冻结保持末值，仅复位沿出 / Fault *)
        ;                                                                      (* 锁存回放（R28） / Replay from latch *)
    ELSE                                                                       (* 非法相位兜底迁安全态 / Illegal phase fallback *)
        _eState := E_DL_BrtState.eFault;                                       (* 迁故障相 / To fault *)
        _bFault := TRUE;                                                       (* 同步锁存 / Latch *)
        _eCause := E_DL_BrtCause.ePhaseBad;                                    (* 成因：非法相位 / Cause: illegal phase *)
END_CASE

(* —— 段 5：出口映射（bError/eState 同源，R191） —— *)
bError := _bFault;                                                             (* 故障标志镜像 / Fault flag mirror *)
eState := _eState;                                                             (* 状态出口 / State outlet *)
eCause := _eCause;                                                             (* 成因出口 / Cause outlet *)
END_FUNCTION_BLOCK

(* ---- FB_DL_BurnerFlameGuard.st ---- *)
(*
  道莅工业代码库 | DL_Device | FB_DL_BurnerFlameGuard
  版本: 1.0.0 | 日期: 2026-11-23 | 轮次: R75
  开源溯源: self-cleanroom（无外部来源；行业池·热工安全通用语义，零代码行复制）
  功能: 燃烧器火焰安全监督——吹扫→点火→火焰建立→运行联锁锁定状态机；点火失败/
        建立失败/运行火焰丢失/联锁丧失均故障锁存并立即关阀，故障相执行安全后吹扫。
  兼容性: CODESYS 3.5 / TwinCAT 3 / 汇川 InoProShop；仅依赖标准 TON / R_TRIG，零厂商私有库
  接口: 输入 bStartCmd/bFlameOk/bInterlockOk/五段定时组态/bReset；输出 bPurgeOut/
        bIgnitionOut/bMainGasOut/bBurnerRun/bSafeShutdown/eState/eCause/bError/nErrId。
        本件无硬件地址依赖，阀与风机输出由上层映射到 %Q。
  码表: 16#0003_031C 故障级：燃烧安全总码（锁存至 bReset 上升沿，归因由 eCause 承载）
        16#0003_040D 信息级：故障相安全后吹扫完成（后吹扫窗到，风机关闭）
        码段说明：0003 段故障子带 03xx / 信息子带 04xx，槽位经全库实扫空闲。
  边界: ① 运行相主燃气阀输出挂 bFlameOk 电平直断——火焰丢失立即关阀，
        锁存经 tFlameLossTol 去抖窗确认（容忍窗内恢复则继续运行）；
        ② 吹扫相检测到火焰信号视作火焰探测器故障（吹扫必须无火）；
        ③ 待机相启动命令而联锁未就绪：拒绝启动（停留在 eIdle），不置故障；
        ④ 六个 TON + 两个 R_TRIG 实例段 0 无条件周期刷新（R7 红线）；
        ⑤ 故障解除唯一路径 = bReset 上升沿 ∧ 组态合法；⑥ 零全局耦合（无 GVL / 无 %I/%Q）。
  邻件比对: registry 扫查 burner/flame 零命中（R75 §3 留痕），无属主。
  修订历史: 2026-11-23 v1.0.0 R75 首版（复杂件批 B1 · C01）
*)

TYPE E_DL_BfgPhase :
(
    eIdle      := 0,   // 待机 | Idle
    ePurge     := 10,  // 前吹扫 | Pre-purge
    eIgnition  := 20,  // 点火试燃 | Ignition trial
    eEstablish := 30,  // 火焰建立确认 | Flame establish confirm
    eRun       := 40,  // 运行联锁锁定 | Run interlocked
    eShutdown  := 50,  // 正常停机后吹扫 | Normal post-purge
    eFault     := 90   // 故障锁存相（含安全后吹扫） | Fault latch phase with post-purge
);
END_TYPE

TYPE E_DL_BfgCause :
(
    eNone          := 0,  // 无故障 | No cause
    eCfgIllegal    := 1,  // 定时组态非法 | Illegal timer configuration
    eInterlock     := 2,  // 联锁条件丧失 | Interlock lost
    eFlameDetPurge := 3,  // 吹扫相火焰信号误现（探测器故障） | Flame signal seen during purge
    eIgnFail       := 4,  // 点火试燃窗内未建立火焰 | No flame in ignition window
    eEstablishFail := 5,  // 建立确认窗内火焰丢失 | Flame lost in establish window
    eFlameLoss     := 6   // 运行相火焰丢失 | Flame loss in run phase
);
END_TYPE

FUNCTION_BLOCK FB_DL_BurnerFlameGuard
VAR_INPUT
    bStartCmd      : BOOL := FALSE;   // 启动命令（电平，自持由上层实现）[-] | Start command level, latching by caller
    bFlameOk       : BOOL := FALSE;   // 火焰检测信号，TRUE=有火 [-] | Flame detector signal, TRUE = flame present
    bInterlockOk   : BOOL := FALSE;   // 联锁总条件（风压/气压/限位外部汇总）[-] | Interlock aggregate from field devices
    tPurgeTime     : TIME := T#60S;   // 前吹扫时长，域 > T#0S | Pre-purge duration
    tIgniteTime    : TIME := T#5S;    // 点火试燃时长，域 > T#0S | Ignition trial duration
    tEstablishTime : TIME := T#10S;   // 火焰建立确认窗，域 > T#0S | Flame establish window
    tPostPurge     : TIME := T#30S;   // 停机/故障后吹扫时长，域 > T#0S | Post-purge duration
    tFlameLossTol  : TIME := T#1S;    // 运行相火焰丢失容忍去抖，域 >= T#0S | Flame loss debounce in run
    bReset         : BOOL := FALSE;   // 复位命令，上升沿清故障 [-] | Reset command, rising edge clears fault
END_VAR
VAR_OUTPUT
    bPurgeOut     : BOOL;              // 吹扫/后吹扫风机输出 [-] | Purge air fan output
    bIgnitionOut  : BOOL;              // 点火输出（火花+引燃气）[-] | Ignition output, spark and pilot
    bMainGasOut   : BOOL;              // 主燃气阀输出（运行相挂火焰信号直断）[-] | Main gas valve output, gated by flame signal
    bBurnerRun    : BOOL;              // 燃烧运行中 [-] | Burner running
    bSafeShutdown : BOOL;              // 安全停机/故障锁存中 [-] | Safe shutdown or fault latched
    eState        : E_DL_BfgPhase;     // 相位出口 | Phase outlet
    eCause        : E_DL_BfgCause;     // 故障成因出口 | Fault cause outlet
    bError        : BOOL;              // 故障锁存标志 [-] | Fault latch flag
    nErrId        : UDINT;             // 事件码，0 = 无事件 | Event code, 0 = none
END_VAR
VAR
    _eState      : E_DL_BfgPhase := E_DL_BfgPhase.eIdle;   // 内部相位（CASE 唯一写入目标） | Internal phase, single write target
    _eCause      : E_DL_BfgCause := E_DL_BfgCause.eNone;   // 故障成因锁存 | Latched fault cause
    _bFault      : BOOL;            // 故障锁存位 | Fault latch bit
    _bPostDone   : BOOL;            // 故障相后吹扫完成保持 | Post-purge done hold in fault phase
    _bCfgBad     : BOOL;            // 组态非法当拍量 [-] | Illegal configuration this scan
    _uInfo       : UDINT;           // 信息码每拍重算 | Info code recomputed per scan
    rtStart      : R_TRIG;          // 启动沿实例，段 0 无条件刷新 | Start edge instance
    rtReset      : R_TRIG;          // 复位沿实例，段 0 无条件刷新 | Reset edge instance
    tonPurge     : TON;             // 前吹扫计时，段 0 无条件刷新 | Pre-purge timer
    tonIgnite    : TON;             // 点火试燃计时，段 0 无条件刷新 | Ignition timer
    tonEstablish : TON;             // 建立确认计时，段 0 无条件刷新 | Establish timer
    tonFlameLoss : TON;             // 运行相火焰丢失去抖，段 0 无条件刷新 | Flame loss debounce timer
    tonPostPurge : TON;             // 后吹扫计时（正常停机与故障相共用），段 0 无条件刷新 | Post-purge timer shared by shutdown and fault
END_VAR

(* —— 段 0：当拍量派生 + 定时器与沿实例无条件周期刷新（R7 红线） —— *)
_bCfgBad := (tPurgeTime <= T#0S) OR (tIgniteTime <= T#0S) OR (tEstablishTime <= T#0S)
         OR (tPostPurge <= T#0S) OR (tFlameLossTol < T#0S);                 // 定时组态域闸 / Timer configuration gate
rtStart(CLK := bStartCmd);                                                  // 启动沿每拍必调 / Start edge every scan
rtReset(CLK := bReset);                                                     // 复位沿每拍必调 / Reset edge every scan
tonPurge(IN := (_eState = E_DL_BfgPhase.ePurge), PT := tPurgeTime);         // 吹扫计时 / Pre-purge timing
tonIgnite(IN := (_eState = E_DL_BfgPhase.eIgnition), PT := tIgniteTime);    // 点火计时 / Ignition timing
tonEstablish(IN := (_eState = E_DL_BfgPhase.eEstablish), PT := tEstablishTime); // 建立计时 / Establish timing
tonFlameLoss(IN := (_eState = E_DL_BfgPhase.eRun) AND (NOT bFlameOk), PT := tFlameLossTol); // 火焰丢失去抖 / Flame loss debounce
tonPostPurge(IN := (_eState = E_DL_BfgPhase.eShutdown) OR (_eState = E_DL_BfgPhase.eFault), PT := tPostPurge); // 后吹扫 / Post-purge timing

(* —— 段 1：单拍量预清零（锁存量不入清单） —— *)
_uInfo := 16#0000_0000;                                                     // 信息码每拍重算 / Info recomputed per scan

(* —— 段 2：复位沿 + 组态域闸 —— *)
IF rtReset.Q AND (NOT _bCfgBad) THEN                                        // 复位沿且组态合法 / Reset edge with legal config
    _bFault    := FALSE;                                                    // 清故障锁存位 / Clear fault latch bit
    _eCause    := E_DL_BfgCause.eNone;                                      // 清成因 / Clear cause
    _bPostDone := FALSE;                                                    // 清后吹扫完成保持 / Clear post-purge hold
    IF _eState = E_DL_BfgPhase.eFault THEN
        _eState := E_DL_BfgPhase.eIdle;                                     // 故障相迁出唯一路径 / Sole exit from fault phase
    END_IF
END_IF
IF _bCfgBad THEN                                                            // 组态域闸 / Configuration gate
    _bFault := TRUE;                                                        // 置故障锁存 / Latch fault
    _eCause := E_DL_BfgCause.eCfgIllegal;                                   // 归因组态非法 / Cause: illegal config
END_IF

(* —— 段 3：相位机（ENUM + CASE，ELSE 兜底） —— *)
CASE _eState OF

E_DL_BfgPhase.eIdle:
    IF rtStart.Q AND bInterlockOk AND (NOT _bFault) THEN
        _eState := E_DL_BfgPhase.ePurge;                                    // 联锁就绪进入前吹扫 / Interlock ready, enter purge
    END_IF                                                                  // 联锁未就绪拒绝启动：停留待机不置故障 / Start refused if interlock not ready

E_DL_BfgPhase.ePurge:
    IF _bFault THEN
        _eState := E_DL_BfgPhase.eFault;                                    // 故障即时迁出 / Leave on fault
    ELSIF NOT bInterlockOk THEN
        _bFault := TRUE;                                                    // 联锁丧失锁存 / Interlock lost latch
        _eCause := E_DL_BfgCause.eInterlock;                                // 归因联锁 / Cause: interlock
        _eState := E_DL_BfgPhase.eFault;
    ELSIF bFlameOk THEN
        _bFault := TRUE;                                                    // 吹扫相见火 = 探测器故障 / Flame in purge = detector fault
        _eCause := E_DL_BfgCause.eFlameDetPurge;                            // 归因探测器 / Cause: flame detector
        _eState := E_DL_BfgPhase.eFault;
    ELSIF tonPurge.Q THEN
        _eState := E_DL_BfgPhase.eIgnition;                                 // 吹扫完成进入点火 / Purge done, ignition trial
    END_IF

E_DL_BfgPhase.eIgnition:
    IF _bFault THEN
        _eState := E_DL_BfgPhase.eFault;                                    // 故障即时迁出 / Leave on fault
    ELSIF NOT bInterlockOk THEN
        _bFault := TRUE;                                                    // 联锁丧失锁存 / Interlock lost latch
        _eCause := E_DL_BfgCause.eInterlock;
        _eState := E_DL_BfgPhase.eFault;
    ELSIF bFlameOk THEN
        _eState := E_DL_BfgPhase.eEstablish;                                // 提前建火提前确认 / Early flame, early establish
    ELSIF tonIgnite.Q THEN
        _bFault := TRUE;                                                    // 点火失败锁存 / Ignition failure latch
        _eCause := E_DL_BfgCause.eIgnFail;                                  // 归因点火 / Cause: ignition fail
        _eState := E_DL_BfgPhase.eFault;
    END_IF

E_DL_BfgPhase.eEstablish:
    IF _bFault THEN
        _eState := E_DL_BfgPhase.eFault;                                    // 故障即时迁出 / Leave on fault
    ELSIF NOT bInterlockOk THEN
        _bFault := TRUE;                                                    // 联锁丧失锁存 / Interlock lost latch
        _eCause := E_DL_BfgCause.eInterlock;
        _eState := E_DL_BfgPhase.eFault;
    ELSIF NOT bFlameOk THEN
        _bFault := TRUE;                                                    // 建立窗内火焰丢失 / Flame lost in establish window
        _eCause := E_DL_BfgCause.eEstablishFail;                            // 归因建立失败 / Cause: establish fail
        _eState := E_DL_BfgPhase.eFault;
    ELSIF tonEstablish.Q THEN
        _eState := E_DL_BfgPhase.eRun;                                      // 火焰稳定进入运行锁定 / Flame stable, run interlocked
    END_IF

E_DL_BfgPhase.eRun:
    IF NOT bInterlockOk THEN
        _bFault := TRUE;                                                    // 运行相联锁丧失立即锁存 / Interlock lost in run, immediate latch
        _eCause := E_DL_BfgCause.eInterlock;
        _eState := E_DL_BfgPhase.eFault;
    ELSIF tonFlameLoss.Q THEN
        _bFault := TRUE;                                                    // 火焰丢失超容忍窗锁存 / Flame loss beyond tolerance latch
        _eCause := E_DL_BfgCause.eFlameLoss;                                // 归因火焰丢失 / Cause: flame loss
        _eState := E_DL_BfgPhase.eFault;
    ELSIF NOT bStartCmd THEN
        _eState := E_DL_BfgPhase.eShutdown;                                 // 正常停机命令进入后吹扫 / Normal stop, post-purge
    END_IF                                                                  // 容忍窗内火焰恢复则继续运行（主燃气阀已挂 bFlameOk 电平） / Recovery inside tolerance keeps running

E_DL_BfgPhase.eShutdown:
    IF tonPostPurge.Q THEN
        _eState := E_DL_BfgPhase.eIdle;                                     // 后吹扫完成回待机 / Post-purge done, back to idle
    END_IF                                                                  // 停机后吹扫期间不判联锁（燃气已关） / Interlock not judged during post-purge, gas closed

E_DL_BfgPhase.eFault:
    IF tonPostPurge.Q AND (NOT _bPostDone) THEN
        _bPostDone := TRUE;                                                 // 故障相后吹扫完成保持 / Post-purge done hold
        _uInfo := 16#0003_040D;                                             // 信息级：安全后吹扫完成 / Info: safe post-purge done
    END_IF                                                                  // 迁出唯一路径 = 段 2 复位沿 / Sole exit is reset edge in segment 2

ELSE
    _bFault := TRUE;                                                        // 非法相位兜底（R6）/ Illegal phase fallback
    _eCause := E_DL_BfgCause.eCfgIllegal;                                   // 归因归并组态 / Cause folded to config
    _eState := E_DL_BfgPhase.eFault;

END_CASE

(* —— 段 4：故障锁存相位迁移闸 —— *)
IF _bFault AND (_eState <> E_DL_BfgPhase.eFault) THEN
    _eState := E_DL_BfgPhase.eFault;                                        // 锁存即入故障相 / Latch enters fault phase
END_IF

(* —— 段 5：出口单点映射（名实同源；安全侧直断） —— *)
bPurgeOut := (_eState = E_DL_BfgPhase.ePurge)
          OR (_eState = E_DL_BfgPhase.eIgnition)
          OR (_eState = E_DL_BfgPhase.eEstablish)
          OR (_eState = E_DL_BfgPhase.eShutdown)
          OR ((_eState = E_DL_BfgPhase.eFault) AND (NOT _bPostDone));       // 风机：吹扫各相 + 故障相未完成段 / Fan in purge phases and unfinished fault purge
bIgnitionOut := ((_eState = E_DL_BfgPhase.eIgnition)
              OR (_eState = E_DL_BfgPhase.eEstablish)) AND (NOT _bFault);   // 点火输出故障即断 / Ignition cut on fault
bMainGasOut := ((_eState = E_DL_BfgPhase.eEstablish)
             OR (_eState = E_DL_BfgPhase.eRun))
             AND (NOT _bFault) AND bFlameOk AND bInterlockOk;               // 主燃气阀挂火焰电平直断（边界①）/ Main gas gated by flame level directly
bBurnerRun := (_eState = E_DL_BfgPhase.eRun) AND (NOT _bFault);             // 运行镜像 / Run mirror
bSafeShutdown := _bFault;                                                   // 安全停机镜像（名实双出口 R191）/ Safe shutdown mirror
eState := _eState;                                                          // 相位出口 / Phase outlet
eCause := _eCause;                                                          // 成因出口 / Cause outlet
bError := _bFault;                                                          // 故障标志同源 / Error flag from latch
IF _bFault THEN
    nErrId := 16#0003_031C;                                                 // 故障锁存码回放 / Replay latched fault code
ELSE
    nErrId := _uInfo;                                                       // 信息码 / Info code
END_IF

END_FUNCTION_BLOCK
